// TwinCAT 3 PLC project PatchPress
// ProgramVersion: 3.1.4026.22
// libraries:
//   Tc2_Standard, * (Beckhoff Automation GmbH)
//   Tc2_System, * (Beckhoff Automation GmbH)
// project tree:
//   DUTs/01_Core/ E_CycleState.TcDUT, E_IndexFault.TcDUT, E_IndexState.TcDUT, E_InitialisingWaitReason.TcDUT, E_MachineState.TcDUT, E_MainDoorLockFault.TcDUT, E_MainDoorLockState.TcDUT, E_OperatorExchangeState.TcDUT, E_OperatorInstruction.TcDUT, E_PartDisposition.TcDUT (not stored), E_ProcessResultCode.TcDUT, E_StoppingWaitReason.TcDUT, E_TablePosition.TcDUT, ST_IndexStatus.TcDUT, ST_MachineCommand.TcDUT, ST_MachineConfig.TcDUT, ST_MachineInputs.TcDUT, ST_MachineOutputs.TcDUT, ST_MachinePermissives.TcDUT, ST_MachineStatus.TcDUT, ST_MainDoorLockStatus.TcDUT, ST_Nest.TcDUT, ST_NestStatistics.TcDUT, ST_OperatorStationStatus.TcDUT, ST_ProcessResult.TcDUT, ST_SafetyStatus.TcDUT (not stored), ST_TestHistory.TcDUT
//   DUTs/01_Core/Machine/ ST_PatchPressInputs.TcDUT, ST_PatchPressOutputs.TcDUT
//   DUTs/02_Components/Motion/ ST_Axis.TcDUT
//   DUTs/04_IO_Mapping/Terminals/ ST_EL3314.TcDUT, ST_EL6633.TcDUT, ST_EK1100.TcDUT (not stored), ST_EL1809.TcDUT (not stored), ST_EL1918.TcDUT, ST_EL2502.TcDUT, ST_EL2809.TcDUT (not stored), ST_EL2904.TcDUT, ST_EL3058.TcDUT, ST_EL3064.TcDUT, ST_EL6070.TcDUT (not stored), ST_EL6652.TcDUT (not stored), ST_EL6910.TcDUT, ST_EL7201.TcDUT, ST_EL9410.TcDUT (not stored), ST_Terminal_Info.TcDUT (not stored)
//   DUTs/07_HMI/ E_LEDs_Mode.TcDUT, E_PLC_Power.TcDUT (not stored), ST_HmiCommands.TcDUT, ST_HmiStatistics.TcDUT, ST_HmiStatus.TcDUT, ST_StatusBanner.TcDUT
//   DUTs/03_Stations/Common/ E_PatchPressStation.TcDUT, E_PatchStationState.TcDUT, ST_PatchStageStatus.TcDUT
//   DUTs/04_IO_Mapping/ ST_PhysicalInputs.TcDUT, ST_PhysicalOutputs.TcDUT
//   DUTs/05_AlarmsAndEvents/ E_AlarmId.TcDUT, E_AlarmSeverity.TcDUT, E_MachineAlarm.TcDUT, ST_ActiveAlarm.TcDUT (not stored), ST_ActiveEvents.TcDUT, ST_AlarmManagerStatus.TcDUT, ST_EVENT.TcDUT, ST_EventsAssigment.TcDUT, ST_EventsAssigmentGeneral.TcDUT (not stored), ST_EventsHistory.TcDUT (not stored), ST_StationEvents.TcDUT
//   GVLs/ GVL_Config.TcGVL, GVL_EtherCAT.TcGVL, GVL_HMI.TcGVL, GVL_IO.TcGVL (not stored), GVL_MASTER.TcGVL, GVL_Motion.TcGVL, GVL_PatchPress_Interface.TcGVL, GVL_Persistent.TcGVL, GVL_Safety.TcGVL
//   / PlcTask.TcTTO
//   POUs/00_Application/ PRG_HmiCommands.TcPOU, PRG_HmiStatus.TcPOU, PRG_Main.TcPOU, PRG_ReadInputs.TcPOU, PRG_WriteOutputs.TcPOU
//   POUs/01_Core/ I_ProcessEquipment.TcIO (not stored)
//   POUs/01_Core/Machine/ FB_IndexedPatchPressMachine.TcPOU, FB_PatchPressCommissioningGuard.TcPOU
//   POUs/01_Core/Process/ FB_ProcessCycle.TcPOU, FB_ProcessStation.TcPOU
//   POUs/02_Components/Door/ FB_MainDoorLock.TcPOU
//   POUs/02_Components/Index/ FB_IndexTable4.TcPOU, FB_NestTableManager.TcPOU, UINT_TO_E_TablePosition.TcPOU
//   POUs/02_Components/Pneumatics/ FB_PuckLocker.TcPOU, FB_Support.TcPOU
//   POUs/03_Stations/HeatStake/ FB_HeatStakeStation.TcPOU
//   POUs/03_Stations/Operator/ FB_OperatorStation.TcPOU
//   POUs/03_Stations/PatchDispense/ FB_PatchDispenseStation.TcPOU
//   POUs/03_Stations/Vision/ FB_VisionStation.TcPOU
//   POUs/04_IO_Mapping/ PRG_TerminalMapping.TcPOU
//   POUs/05_AlarmsAndEvents/ FB_EventsManager.TcPOU, PRG_Events.TcPOU
//   POUs/06_Utilities/ FB_TerminalInfo.TcPOU (not stored), F_ScaleLinear.TcPOU
//   POUs/ MAIN.TcPOU
// real-time tasks:
//   TASK PlcTask: cycle T#10ms, priority 20, ADS port 350
// motion (NC):
//   TASK NC-Task 1 SAF: cycle T#2ms, priority 4, ADS port 501
//   TASK NC-Task 1 SVB: cycle T#10ms, priority 8, ADS port 511
//   AXIS M1 (id 1)
//     OtherSettings: AllowMotionCmdToSlave=true
//     encoder EncType=19
//       EncPara: MaxCount=#xffffffff
//     drive DrvType=16
//       DrvPara: MaxCount=#xffffffff, DriveControlDWord=#x00020000
//         Analog: TorqueSetpointScale=10, ScaleFactorActTorque=0.1
//         TimeComp: TaskDelayCycles=1
//     controller CtrType=1
//       CtrPara: PriorControlFactor=1
//         Observer: BandWidth=20
//   AXIS M2 (id 2)
//     OtherSettings: AllowMotionCmdToSlave=true
//     encoder EncType=19
//       EncPara: MaxCount=#xffffffff
//     drive DrvType=16
//       DrvPara: MaxCount=#xffffffff, DriveControlDWord=#x00020000
//         Analog: TorqueSetpointScale=10, ScaleFactorActTorque=0.1
//         TimeComp: TaskDelayCycles=1
//     controller CtrType=1
//       CtrPara: PriorControlFactor=1
//         Observer: BandWidth=20
//   AXIS M3 (id 3)
//     OtherSettings: AllowMotionCmdToSlave=true
//     encoder EncType=19
//       EncPara: MaxCount=#xffffffff
//     drive DrvType=16
//       DrvPara: MaxCount=#xffffffff, DriveControlDWord=#x00020000
//         Analog: TorqueSetpointScale=10, ScaleFactorActTorque=0.1
//         TimeComp: TaskDelayCycles=1
//     controller CtrType=1
//       CtrPara: PriorControlFactor=1
//         Observer: BandWidth=20
// I/O:
//   DEVICE Device 1 (EtherCAT), AmsNetId 172.18.239.27.2.1
//     Term 1 (EK1100) [EK1100 EtherCAT Coupler (2A E-Bus)]
//       Term 2 (EL6070-0033) [EL6070-0033 1Ch. Licence key terminal, individual licences]
//       Term 3 (EL6910) [EL6910, TwinSAFE PLC]
//       Term 4 (EL1918) [EL1918, 8Ch. Safety Input 24V, TwinSAFE]
//         modules: Module 1 (FSOE), Module 2 (FSLOGIC)
//       Term 5 (EL1918) [EL1918, 8Ch. Safety Input 24V, TwinSAFE]
//         modules: Module 1 (FSOE), Module 2 (FSLOGIC)
//       Term 6 (EL2904) [EL2904, 4 Ch. Safety Output 24V, 0.5A, TwinSAFE]
//         modules: Module 1 (FSOES), Module 2 (DO)
//       Term 7 (EL1809) [EL1809 16Ch. Dig. Input 24V, 3ms]
//       Term 8 (EL1809) [EL1809 16Ch. Dig. Input 24V, 3ms]
//       Term 9 (EL2809-0015) [EL2809-0015 16Ch. Dig. Output 24V DC, 0.35A, not short-circuit proof]
//       Term 10 (EL2809-0015) [EL2809-0015 16Ch. Dig. Output 24V DC, 0.35A, not short-circuit proof]
//       Term 11 (EL3058) [EL3058 8Ch. Ana. Input 4-20mA]
//       Term 12 (EL9410) [EL9410 E-Bus Power Supplier  (Diagnostics)]
//       Term 13 (EL2502) [EL2502 2Ch. PWM output, 24V]
//       Term 14 (EL9576) [EL9576 Brake chopper terminal]
//       Term 15 (EL7201-9014) [EL7201-9014 1Ch. MDP742 Servo motor output stage with OCT (50V, 2.8A RMS) and STO input]
//       Term 16 (EL7201-9014) [EL7201-9014 1Ch. MDP742 Servo motor output stage with OCT (50V, 2.8A RMS) and STO input]
//       Term 17 (EL7201-9014) [EL7201-9014 1Ch. MDP742 Servo motor output stage with OCT (50V, 2.8A RMS) and STO input]
//       Term 18 (EL2904) [EL2904, 4 Ch. Safety Output 24V, 0.5A, TwinSAFE]
//         modules: Module 1 (FSOES), Module 2 (DO)
//       Term 19 (EL1809) [EL1809 16Ch. Dig. Input 24V, 3ms]
//       Term 20 (EL3314-0092) [EL3314-0092 4Ch. Ana Input Thermocouple (TC), TwinSAFE SC]
//       Term 21 (EL6633) [EL6633 PROFINET IO Controller]
//       Term 23 (EL9011) [EL9011 End Terminal]
//     Box 22 (VABX-A-S-EL-E12-CTED-ECM12) [VABX-A-S-EL-E12-CTED-ECM12] (disabled)
// variable links:
//   Device 1 (EtherCAT) <-> Device 1 (EtherCAT)/Term 1 (EK1100)/Term 3 (EL6910)
//     Term 1 (EK1100)/Term 18 (EL2904)/Module 1 (FSOES)/RxPDO/FSOE <-> ConnectionInputs/TwinSafeGroup1.Term 18 (EL2904) - Module 1 (FSOES)_6 TxPDO
//     Term 1 (EK1100)/Term 6 (EL2904)/Module 1 (FSOES)/RxPDO/FSOE <-> ConnectionInputs/TwinSafeGroup1.Term 6 (EL2904) - Module 1 (FSOES)_5 TxPDO
//     Term 1 (EK1100)/Term 18 (EL2904)/Module 1 (FSOES)/TxPDO/FSOE <-> ConnectionOutputs/TwinSafeGroup1.Term 18 (EL2904) - Module 1 (FSOES)_6 RxPDO
//     Term 1 (EK1100)/Term 6 (EL2904)/Module 1 (FSOES)/TxPDO/FSOE <-> ConnectionOutputs/TwinSafeGroup1.Term 6 (EL2904) - Module 1 (FSOES)_5 RxPDO
//     Term 1 (EK1100)/Term 4 (EL1918)/Module 1 (FSOE)/FSoE Inputs/FSOE <-> ConnectionOutputs/TwinSafeGroup1.Term 4 (EL1918) - Module 1 (FSOE)_3 RxPDO
//     Term 1 (EK1100)/Term 5 (EL1918)/Module 1 (FSOE)/FSoE Inputs/FSOE <-> ConnectionOutputs/TwinSafeGroup1.Term 5 (EL1918) - Module 1 (FSOE)_4 RxPDO
//     Term 1 (EK1100)/Term 4 (EL1918)/Module 1 (FSOE)/FSoE Outputs/FSOE <-> ConnectionInputs/TwinSafeGroup1.Term 4 (EL1918) - Module 1 (FSOE)_3 TxPDO
//     Term 1 (EK1100)/Term 5 (EL1918)/Module 1 (FSOE)/FSoE Outputs/FSOE <-> ConnectionInputs/TwinSafeGroup1.Term 5 (EL1918) - Module 1 (FSOE)_4 TxPDO
//   NC-Task 1 SAF/Axes/M1 <-> Device 1 (EtherCAT)/Term 1 (EK1100)/Term 15 (EL7201-9014)
//     Drive/Inputs/In/nDcOutputTime <-> InfoData/DcOutputShift
//     Drive/Inputs/In/nState1 <-> DRV Statusword/Statusword
//     Drive/Inputs/In/nState2 <-> DRV Statusword/Statusword @bit 8
//     Drive/Inputs/In/nState4 @bit 1 <-> WcState/InputToggle
//     Drive/Inputs/In/nState4 <-> WcState/WcState
//     Drive/Outputs/Out/nCtrl1 <-> DRV Controlword/Controlword
//     Drive/Outputs/Out/nCtrl2 <-> DRV Controlword/Controlword @bit 8
//     Drive/Outputs/Out/nDataOut2 <-> DRV Target velocity/Target velocity
//     Enc/Inputs/In/nDataIn1 <-> FB Position/Position
//     Enc/Inputs/In/nDcInputTime <-> InfoData/DcInputShift
//     Enc/Inputs/In/nState4 @bit 1 <-> WcState/InputToggle
//     Enc/Inputs/In/nState4 <-> WcState/WcState
//   NC-Task 1 SAF/Axes/M2 <-> Device 1 (EtherCAT)/Term 1 (EK1100)/Term 16 (EL7201-9014)
//     Drive/Inputs/In/nDcOutputTime <-> InfoData/DcOutputShift
//     Drive/Inputs/In/nState1 <-> DRV Statusword/Statusword
//     Drive/Inputs/In/nState2 <-> DRV Statusword/Statusword @bit 8
//     Drive/Inputs/In/nState4 @bit 1 <-> WcState/InputToggle
//     Drive/Inputs/In/nState4 <-> WcState/WcState
//     Drive/Outputs/Out/nCtrl1 <-> DRV Controlword/Controlword
//     Drive/Outputs/Out/nCtrl2 <-> DRV Controlword/Controlword @bit 8
//     Drive/Outputs/Out/nDataOut2 <-> DRV Target velocity/Target velocity
//     Enc/Inputs/In/nDataIn1 <-> FB Position/Position
//     Enc/Inputs/In/nDcInputTime <-> InfoData/DcInputShift
//     Enc/Inputs/In/nState4 @bit 1 <-> WcState/InputToggle
//     Enc/Inputs/In/nState4 <-> WcState/WcState
//   NC-Task 1 SAF/Axes/M3 <-> Device 1 (EtherCAT)/Term 1 (EK1100)/Term 17 (EL7201-9014)
//     Drive/Inputs/In/nDcOutputTime <-> InfoData/DcOutputShift
//     Drive/Inputs/In/nState1 <-> DRV Statusword/Statusword
//     Drive/Inputs/In/nState2 <-> DRV Statusword/Statusword @bit 8
//     Drive/Inputs/In/nState4 @bit 1 <-> WcState/InputToggle
//     Drive/Inputs/In/nState4 <-> WcState/WcState
//     Drive/Outputs/Out/nCtrl1 <-> DRV Controlword/Controlword
//     Drive/Outputs/Out/nCtrl2 <-> DRV Controlword/Controlword @bit 8
//     Drive/Outputs/Out/nDataOut2 <-> DRV Target velocity/Target velocity
//     Enc/Inputs/In/nDataIn1 <-> FB Position/Position
//     Enc/Inputs/In/nDcInputTime <-> InfoData/DcInputShift
//     Enc/Inputs/In/nState4 @bit 1 <-> WcState/InputToggle
//     Enc/Inputs/In/nState4 <-> WcState/WcState
//   PatchPress/PatchPress Instance <-> Device 1 (EtherCAT)/Term 1 (EK1100)/Term 10 (EL2809-0015)
//     PlcTask Inputs/GVL_EtherCAT.stTerm10_EL2809.stTerminalInfo.nTerminal_State <-> InfoData/State
//     PlcTask Outputs/GVL_EtherCAT.stTerm10_EL2809.iEL2809_Ch{1..16} <-> Channel {1..16}/Output  (16 links)
//   PatchPress/PatchPress Instance <-> Device 1 (EtherCAT)/Term 1 (EK1100)/Term 11 (EL3058)
//     PlcTask Inputs/GVL_EtherCAT.stTerm11_EL3058.iEL3058_Ch{1..8} <-> AI Standard Channel {1..8}/Value  (8 links)
//     PlcTask Inputs/GVL_EtherCAT.stTerm11_EL3058.stTerminalInfo.nTerminal_State <-> InfoData/State
//   PatchPress/PatchPress Instance <-> Device 1 (EtherCAT)/Term 1 (EK1100)/Term 19 (EL1809)
//     PlcTask Inputs/GVL_EtherCAT.stTerm19_EL1809.iEL1809_Ch{1..16} <-> Channel {1..16}/Input  (16 links)
//     PlcTask Inputs/GVL_EtherCAT.stTerm19_EL1809.stTerminalInfo.nTerminal_State <-> InfoData/State
//   PatchPress/PatchPress Instance <-> Device 1 (EtherCAT)/Term 1 (EK1100)/Term 3 (EL6910)
//     PlcTask Inputs/GVL_Safety.bMainDoorClosed <-> StandardInputs/Standard Out Var 8
//     PlcTask Inputs/GVL_Safety.bMainDoorLocked <-> StandardInputs/Standard Out Var 9
//     PlcTask Inputs/GVL_Safety.bMainDoorUnSafe <-> StandardInputs/Standard Out Var 10
//     PlcTask Inputs/GVL_Safety.bResetButtonPressed <-> StandardInputs/Standard Out Var 7
//     PlcTask Inputs/GVL_Safety.bSafetyOk <-> StandardInputs/Standard Out Var 12
//     PlcTask Inputs/GVL_Safety.bTwoHandSafe <-> StandardInputs/Standard Out Var 16
//     PlcTask Outputs/GVL_IO.stOutputs/bAirSupplyEnable <-> StandardOutputs/Standard In Var 11
//     PlcTask Outputs/GVL_IO.stOutputs/bMainDoorLockRequest <-> StandardOutputs/Standard In Var 14
//     PlcTask Outputs/GVL_IO.stOutputs/bSafetyErrorAcknowledgementRequest <-> StandardOutputs/Standard In Var 1
//     PlcTask Outputs/GVL_IO.stOutputs/bSafetyRunRequest <-> StandardOutputs/Standard In Var 15
//   PatchPress/PatchPress Instance <-> Device 1 (EtherCAT)/Term 1 (EK1100)/Term 7 (EL1809)
//     PlcTask Inputs/GVL_EtherCAT.stTerm7_EL1809.iEL1809_Ch{1..16} <-> Channel {1..16}/Input  (16 links)
//     PlcTask Inputs/GVL_EtherCAT.stTerm7_EL1809.stTerminalInfo.nTerminal_State <-> InfoData/State
//   PatchPress/PatchPress Instance <-> Device 1 (EtherCAT)/Term 1 (EK1100)/Term 8 (EL1809)
//     PlcTask Inputs/GVL_EtherCAT.stTerm8_EL1809.iEL1809_Ch{1..16} <-> Channel {1..16}/Input  (16 links)
//     PlcTask Inputs/GVL_EtherCAT.stTerm8_EL1809.stTerminalInfo.nTerminal_State <-> InfoData/State
//   PatchPress/PatchPress Instance <-> Device 1 (EtherCAT)/Term 1 (EK1100)/Term 9 (EL2809-0015)
//     PlcTask Inputs/GVL_EtherCAT.stTerm9_EL2809.stTerminalInfo.nTerminal_State <-> InfoData/State
//     PlcTask Outputs/GVL_EtherCAT.stTerm9_EL2809.iEL2809_Ch{1..16} <-> Channel {1..16}/Output  (16 links)

CONFIGURATION PatchPress
    RESOURCE PLC ON TwinCAT3
        TASK PlcTask(INTERVAL := T#10ms, PRIORITY := 20);
        PROGRAM MAIN WITH PlcTask : MAIN;
    END_RESOURCE
END_CONFIGURATION

// ---- DUTs/01_Core/E_CycleState.TcDUT
{attribute 'qualified_only'}
{attribute 'strict'}
{attribute 'to_string'}
TYPE E_CycleState :
(
    // CYCLE INITIALISATION
    Disabled                        := 0,
    Initialising                    := 10,
    WaitingForProcessCycleTrigger   := 20,
	
    // INDEX POSITION RECOVERY
    EvaluatingIndexPosition         := 30,
    RequestingIndexPositionRecovery := 40,
    WaitingForIndexPositionRecovery := 50,

    // INDEX MOVEMENT
    ValidatingIndexPermissives      := 60,
    RequestingIndexMove             := 70,
    WaitingForIndexStart            := 80,
    WaitingForIndexComplete         := 90,

    // NEST AND PROCESS PREPARATION
    UpdatingNestPositions           := 100,
    EvaluatingProcessNest           := 110,
    SkippingProcessNest             := 120,

    // SUPPORT EXTENSION
    RequestingSupportsExtend        := 130,
    WaitingForSupportsExtended      := 140,

    // PROCESS EXECUTION
    PreparingProcessStations        := 150,
    WaitingForProcessStationsReady  := 160,
    StartingProcesses               := 170,
    WaitingForProcessesRunning      := 180,
    WaitingForProcessesComplete     := 190,

    // PROCESS RESULT
    CapturingProcessResult          := 200,
    StoringProcessResult            := 210,

    // SUPPORT RETRACTION
    RequestingSupportsRetract       := 220,
    WaitingForSupportsRetracted     := 230,

    // OPERATOR EXCHANGE
    PreparingOperatorExchange       := 240,
    WaitingForOperatorExchange      := 250,
    ConfirmingOperatorExchange      := 260,

    // CYCLE COMPLETION
    CycleComplete                   := 270,

    // TERMINAL STATES
    ControlledStop                  := 900,
    Fault                           := 999
);
END_TYPE

// ---- DUTs/01_Core/E_IndexFault.TcDUT
{attribute 'qualified_only'}
{attribute 'strict'}
{attribute 'to_string'}
TYPE E_IndexFault :
(
    None := 0,
    InitialPositionInvalid,
    SupportRetractTimeout,
    RotationTimeout,
    StopAndLockTimeout,
    PositionInvalid,
    SupportExtendTimeout,
    TwoHandReleasedDuringMovement,
    WrongPositionTimeout,
    SafetyLostDuringMovement,
    MovementPermissiveLost
);
END_TYPE

// ---- DUTs/01_Core/E_IndexState.TcDUT
{attribute 'qualified_only'}
{attribute 'strict'}
{attribute 'to_string'}
TYPE E_IndexState :
(
    Disabled := 0,
    Initialising,
    Idle,
    RetractingSupport,
    WaitingSupportRetracted,
    RotatingPortA,
    WrongPositionRecovery,
    StoppingPortB,
    VerifyingPosition,
    ExtendingSupport,
    WaitingSupportExtended,
    ProcessPositionReady,
    WaitingOperatorExchange,
    Complete,
    Stopping,
    Fault
);
END_TYPE

// ---- DUTs/01_Core/E_InitialisingWaitReason.TcDUT
{attribute 'qualified_only'}
{attribute 'strict'}
{attribute 'to_string'}
TYPE E_InitialisingWaitReason :
(
    None := 0,
    SafetyNotReady := 10,
    FsoeNotReady := 20,
    SafetyLogicNotReady := 30,
    AirSupplyNotReady := 40,
    MainDoorNotReady := 50,
    IndexNotReady := 60,
    StationsNotHome := 70
);
END_TYPE

// ---- DUTs/01_Core/E_MachineState.TcDUT
{attribute 'qualified_only'}
{attribute 'strict'}
{attribute 'to_string'}
TYPE E_MachineState :
(
    PowerUp      := 0,
    Fault        := 1,
    Stopping     := 2,
    Stopped      := 3,
    Initialising := 4,
    ReadyToStart := 5,
    AutoCycle    := 6,
    Manual       := 7
);
END_TYPE

// ---- DUTs/01_Core/E_MainDoorLockFault.TcDUT
{attribute 'qualified_only'}
{attribute 'strict'}
{attribute 'to_string'}
TYPE E_MainDoorLockFault :
(
    None := 0,
    LockTimeout := 10,
    UnlockTimeout := 20,
    DoorNotClosed := 30,
    FeedbackMismatch := 40
);
END_TYPE

// ---- DUTs/01_Core/E_MainDoorLockState.TcDUT
{attribute 'qualified_only'}
{attribute 'strict'}
{attribute 'to_string'}
TYPE E_MainDoorLockState :
(
    Disabled := 0,
    Unlocked := 10,
    Locking := 20,
    Locked := 30,
    Unlocking := 40,
    Fault := 999
);
END_TYPE

// ---- DUTs/01_Core/E_OperatorExchangeState.TcDUT
{attribute 'qualified_only'}
{attribute 'strict'}
{attribute 'to_string'}
TYPE E_OperatorExchangeState :
(
    Idle := 0,
    EvaluateNest := 10,
    WaitingForPartRemoval := 20,
    WaitingForRejectConfirmation := 30,
    WaitingForPuckRemoval := 40,
    WaitingForNewPuck := 50,
    WaitingForPuckLocked := 60,
    WaitingForPartLoading := 70,
    ExchangeComplete := 80,
    WaitingForTableIndexComplete := 90,
    Fault := 999
);
END_TYPE

// ---- DUTs/01_Core/E_OperatorInstruction.TcDUT
{attribute 'qualified_only'}
{attribute 'strict'}
{attribute 'to_string'}
TYPE E_OperatorInstruction :
(
    None := 0,
    LoadInitialPuck := 10,
    WaitPuckLocking := 20,
    RemovePassedPart := 30,
    RemoveFailedPart := 40,
    PlacePartInRejectBin := 50,
    RemoveReleasedPuck := 60,
    LoadNewPuck := 70,
    LoadPart := 80,
    ReadyToIndex := 90,
    ReadyToIndexEmpty := 100,
    TableIndexing := 110,
    RestoreUnexpectedlyRemovedPuck := 120
);
END_TYPE

// ---- DUTs/01_Core/E_ProcessResultCode.TcDUT
{attribute 'qualified_only'}
{attribute 'strict'}
{attribute 'to_string'}
TYPE E_ProcessResultCode :
(
	None := 0,
    Pass,
    Fail,
    Aborted,
    EquipmentFault,
    CommunicationFault,
    Timeout
);
END_TYPE

// ---- DUTs/01_Core/E_StoppingWaitReason.TcDUT
{attribute 'qualified_only'}
{attribute 'strict'}
{attribute 'to_string'}
TYPE E_StoppingWaitReason :
(
    None := 0,
    IndexStillMoving := 10,
    MainDoorTransition := 20
);
END_TYPE

// ---- DUTs/01_Core/E_TablePosition.TcDUT
{attribute 'qualified_only'}
{attribute 'strict'}
{attribute 'to_string'}
TYPE E_TablePosition :
(
	Unknown := 0,
    Position1 := 1,
    Position2 := 2,
    Position3 := 3,
    Position4 := 4
);
END_TYPE

// ---- DUTs/01_Core/Machine/ST_PatchPressInputs.TcDUT
TYPE ST_PatchPressInputs :
STRUCT
    // EPLAN Term 7 - EL1809
    b48VPowerSupplyOk                   : BOOL;
    bLoadingStationEaglePresent         : BOOL;
    bRejectChutePartPresent             : BOOL;
    bHeatStakeEagleAssemblyPresent      : BOOL;
    bHeatStakePatchPresent              : BOOL;
    bPbupMagnetPresent                  : BOOL;

    // EPLAN Term 8 - EL1809
    bStation1SupportRetracted           : BOOL;
    bStation1SupportExtended            : BOOL;
    bStation2SupportRetracted           : BOOL;
    bStation2SupportExtended            : BOOL;
    bStation3SupportRetracted           : BOOL;
    bStation3SupportExtended            : BOOL;
    bHorizontalMiniSlideRetracted       : BOOL;
    bHorizontalMiniSlideExtended        : BOOL;
    bVerticalMiniSlideRetracted         : BOOL;
    bVerticalMiniSlideExtended          : BOOL;
    bIntermediateModuleRetracted        : BOOL;
    bIntermediateModuleExtended         : BOOL;
    bRotaryGripperOpened                : BOOL;
    bRotaryGripperClosed                : BOOL;
    bRotaryGripperPick0                 : BOOL;
    bRotaryGripperPlace180              : BOOL;

    // EPLAN Term 19 - EL1809
    bMembraneTransferRetracted          : BOOL;
    bMembraneTransferExtended           : BOOL;
    bMiddleRockerDown                   : BOOL;
    bMiddleRockerUp                     : BOOL;
    bBottomRockerDown                   : BOOL;
    bBottomRockerUp                     : BOOL;
    bTopRockerDown                      : BOOL;
    bTopRockerUp                        : BOOL;

    // EPLAN Term 11 / 20
    iMainAirPressureRaw                 : INT;
    iProportionalPressureActualRaw      : INT;
    iCartridgeHeater1TemperatureRaw     : INT;
    iCartridgeHeater2TemperatureRaw     : INT;
    iOverTemperatureRaw                 : INT;
END_STRUCT
END_TYPE

// ---- DUTs/01_Core/Machine/ST_PatchPressOutputs.TcDUT
TYPE ST_PatchPressOutputs :
STRUCT
    // Pneumatic commands are logical commands only at this stage.
    // Physical Festo manifold PDO mapping must be created after the manifold scan.
    bStation1SupportExtend              : BOOL;
    bStation1SupportRetract             : BOOL;
    bStation2SupportExtend              : BOOL;
    bStation2SupportRetract             : BOOL;
    bStation3SupportExtend              : BOOL;
    bStation3SupportRetract             : BOOL;
    bHorizontalMiniSlideExtend          : BOOL;
    bHorizontalMiniSlideRetract         : BOOL;
    bVerticalMiniSlideExtend            : BOOL;
    bVerticalMiniSlideRetract           : BOOL;
    bIntermediateModuleExtend           : BOOL;
    bIntermediateModuleRetract          : BOOL;
    bRotaryGripperOpen                  : BOOL;
    bRotaryGripperClose                 : BOOL;
    bRotaryGripperPick0                 : BOOL;
    bRotaryGripperPlace180              : BOOL;
    bMembraneTransferExtend             : BOOL;
    bMembraneTransferRetract            : BOOL;
    bMiddleRockerDown                   : BOOL;
    bMiddleRockerUp                     : BOOL;
    bBottomRockerDown                   : BOOL;
    bBottomRockerUp                     : BOOL;
    bTopRockerDown                      : BOOL;
    bTopRockerUp                        : BOOL;

    // Heater / pressure logical commands.
    rHeater1DutyPercent                 : REAL;
    rHeater2DutyPercent                 : REAL;
    rPressureSetpointBar                : REAL;
END_STRUCT
END_TYPE

// ---- DUTs/01_Core/ST_IndexStatus.TcDUT
TYPE ST_IndexStatus :
STRUCT
    eState                    : E_IndexState;
    eFault                    : E_IndexFault;
    eCurrentPosition          : E_TablePosition;

    bReady                    : BOOL;
    bBusy                     : BOOL;
    bFaulted                  : BOOL;
    bDonePulse                : BOOL;

    bManualMoveActive         : BOOL;
    bPositionRecoveryActive   : BOOL;
    bSamePositionDetected     : BOOL;
    bWrongPositionTimerActive : BOOL;
    bTwoHandRequired          : BOOL;

    bProcessPositionReady     : BOOL;
    bWaitingOperatorExchange  : BOOL;

    bSupportRetracted         : BOOL;
    bSupportExtended          : BOOL;
    bTableReady               : BOOL;
    bTableLocked              : BOOL;
	
END_STRUCT
END_TYPE

// ---- DUTs/01_Core/ST_MachineCommand.TcDUT
TYPE ST_MachineCommand :
STRUCT
    bStart                : BOOL;
    bStop                 : BOOL;
    bReset                : BOOL;
    bManualRequest        : BOOL;
    bManualIndexForward   : BOOL;
    bManualIndexHome      : BOOL;
    bIndexerManualEnable  : BOOL;
    bManualMainDoorUnlock : BOOL;
    bAcknowledge          : BOOL;
    bAcknowledgePuckRemovalFault : BOOL;
    uiResetStatisticsNestId : UINT;
END_STRUCT
END_TYPE

// ---- DUTs/01_Core/ST_MachineConfig.TcDUT
TYPE ST_MachineConfig :
STRUCT
    tInitialiseTimeout       : TIME := T#20S;
    tStoppingTimeout         : TIME := T#15S;
    tIndexTimeout            : TIME := T#10S;
    tIndexRotateDelay        : TIME := T#500MS;
    tIndexStopDelay          : TIME := T#1S;
    tIndexSupportTimeout     : TIME := T#5S;
    tTwoHandHold             : TIME := T#500MS;
    tTwoHandRecoveryTimeout  : TIME := T#10S;
    tDoorLockTimeout         : TIME := T#10S;
    tDoorUnlockTimeout       : TIME := T#10S;
    tOperatorIdleTimeout     : TIME := T#30S;
    eOperatorPosition        : E_TablePosition := E_TablePosition.Position1;
    ePatchDispensePosition   : E_TablePosition := E_TablePosition.Position2;
    eHeatStakePosition       : E_TablePosition := E_TablePosition.Position3;
    eVisionPosition          : E_TablePosition := E_TablePosition.Position4;
    eRejectPosition          : E_TablePosition := E_TablePosition.Position1;
    bRequireTwoHandsForIndex : BOOL := TRUE;
    bAllowEmptyNestIndex     : BOOL := TRUE;
    bRequireRejectConfirm    : BOOL := TRUE;
    aNestEnabled             : ARRAY[1..4] OF BOOL := [TRUE, TRUE, TRUE, TRUE];
END_STRUCT
END_TYPE

// ---- DUTs/01_Core/ST_MachineInputs.TcDUT
TYPE ST_MachineInputs :
STRUCT
    bStartButton                  : BOOL;
    bStopButton                   : BOOL;
    bResetButton                  : BOOL;
    bTwoHandsSafe                 : BOOL;
    bTouchButtonLeft              : BOOL;
    bTouchButtonRight             : BOOL;
    bUp24VPowerSupplyOk           : BOOL;
    bUs24VPowerSupplyOk           : BOOL;
    b48VPowerSupplyOk             : BOOL;
    bEmergencyStopChannel1        : BOOL;
    bEmergencyStopChannel2        : BOOL;
    bMainDoorChannel1             : BOOL;
    bMainDoorChannel2             : BOOL;
    bMainDoorFeedback             : BOOL;
    bLeftFlapChannel1             : BOOL;
    bLeftFlapChannel2             : BOOL;
    bRightFlapChannel1            : BOOL;
    bRightFlapChannel2            : BOOL;
    bMainDoorClosed               : BOOL;
    bMainDoorLocked               : BOOL;
    bMainDoorUnsafe               : BOOL;
    bMainDoorDiagnosticOk         : BOOL;
    bMs6FeedbackOk                : BOOL;
    bAirExhausted                 : BOOL;
    stSafety                      : ST_SafetyStatus;
    bEventFault                   : BOOL;
    bEventCycleStopRequest        : BOOL;
    bIndexReady                   : BOOL;
    bIndexLocked                  : BOOL;
    bIndexCompletedSensor         : BOOL;
    eIndexPosition                : E_TablePosition;
    bLoadingStationEaglePresent   : BOOL;
    bRejectChutePartPresent       : BOOL;
    bHeatStakeEaglePresent        : BOOL;
    bHeatStakePatchPresent        : BOOL;
    bPbupMagnetPresent            : BOOL;
    bStation1SupportRetracted     : BOOL;
    bStation1SupportExtended      : BOOL;
    bStation2SupportRetracted     : BOOL;
    bStation2SupportExtended      : BOOL;
    bStation3SupportRetracted     : BOOL;
    bStation3SupportExtended      : BOOL;
    bHorizontalMiniSlideRetracted : BOOL;
    bHorizontalMiniSlideExtended  : BOOL;
    bVerticalMiniSlideRetracted   : BOOL;
    bVerticalMiniSlideExtended    : BOOL;
    bIntermediateModuleRetracted  : BOOL;
    bIntermediateModuleExtended   : BOOL;
    bRotaryGripperOpened          : BOOL;
    bRotaryGripperClosed          : BOOL;
    bRotaryGripperPick0           : BOOL;
    bRotaryGripperPlace180        : BOOL;
    bMembraneTransferRetracted    : BOOL;
    bMembraneTransferExtended     : BOOL;
    bMiddleRockerDown             : BOOL;
    bMiddleRockerUp               : BOOL;
    bBottomRockerDown             : BOOL;
    bBottomRockerUp               : BOOL;
    bTopRockerDown                : BOOL;
    bTopRockerUp                  : BOOL;
    uiMainAirPressureRaw          : UINT;
    uiPressureRegulatorActualRaw  : UINT;
END_STRUCT
END_TYPE

// ---- DUTs/01_Core/ST_MachineOutputs.TcDUT
TYPE ST_MachineOutputs :
STRUCT
    bSafetyRunRequest                  : BOOL;
    bSafetyResetRequest                : BOOL;
    bSafetyErrorAcknowledgementRequest : BOOL;
    bAirSupplyEnable                   : BOOL;
    bMainDoorLockRequest               : BOOL;
    bIndexRotatePortA                  : BOOL;
    bIndexStopPortB                    : BOOL;
    bIndexSupportExtend                : BOOL;
    bIndexSupportRetract               : BOOL;
    bLedStart                          : BOOL;
    bLedReset                          : BOOL;
    bLedPass                           : BOOL;
    bLedFail                           : BOOL;
    bInternalLight                     : BOOL;
    bNestLight                         : BOOL;
END_STRUCT
END_TYPE

// ---- DUTs/01_Core/ST_MachinePermissives.TcDUT
TYPE ST_MachinePermissives :
STRUCT
    bSafetyIndexPermissive   : BOOL;
    bOperatorIndexPermissive : BOOL;
    bStationsIndexPermissive : BOOL;
    bIndexMoveAllowed        : BOOL;
    bAirSupplyReady          : BOOL;
    bDoorInitialisationReady : BOOL;
    bIndexInitialisationReady: BOOL;
    bStationsHome            : BOOL;
    bInitialisationAllowed   : BOOL;
    bAutoCycleAllowed        : BOOL;
END_STRUCT
END_TYPE

// ---- DUTs/01_Core/ST_MachineStatus.TcDUT
TYPE ST_MachineStatus :
STRUCT
    eMachineState           : E_MachineState;
    eIndexState             : E_IndexState;
    stIndexStatus           : ST_IndexStatus;
    stMainDoorLock          : ST_MainDoorLockStatus;
    eInitialisingWaitReason : E_InitialisingWaitReason;
    eStoppingWaitReason     : E_StoppingWaitReason;
    eOperatorExchangeState  : E_OperatorExchangeState;
    eOperatorInstruction    : E_OperatorInstruction;
    stOperatorStation       : ST_OperatorStationStatus;
    stPatchDispense         : ST_PatchStageStatus;
    stHeatStake             : ST_PatchStageStatus;
    stVision                : ST_PatchStageStatus;
    bReady                  : BOOL;
    bBusy                   : BOOL;
    bFaulted                : BOOL;
    bInitialisationTimeoutFault : BOOL;
    bStoppingTimeoutFault   : BOOL;
    bSafetyStopRequested    : BOOL;
    bSafetyRunRequested     : BOOL;
    bEventFault             : BOOL;
    bCycleStopRequested     : BOOL;
    bIndexPermissive        : BOOL;
    bEnableSetting          : BOOL;
    bAllStationsCommissioned: BOOL;
    bAutoCycleAllowed       : BOOL;
    stPermissives           : ST_MachinePermissives;
    stLastResult            : ST_ProcessResult;
    aNest                   : ARRAY[1..4] OF ST_Nest;
    aNestStatistics         : ARRAY[1..4] OF ST_NestStatistics;
    sMachineMessage         : STRING(160);
    sOperatorMessage        : STRING(255);
    sAutoCycleBlockReason   : STRING(160);
END_STRUCT
END_TYPE

// ---- DUTs/01_Core/ST_MainDoorLockStatus.TcDUT
TYPE ST_MainDoorLockStatus :
STRUCT
    eState                  : E_MainDoorLockState;
    eFault                  : E_MainDoorLockFault;
    bDoorClosed             : BOOL;
    bDoorLocked             : BOOL;
    bDoorUnsafe             : BOOL;
    bLockRequest            : BOOL;
    bLockOutput             : BOOL;
    bReadyForAutomatic      : BOOL;
    bUnlockPermissive       : BOOL;
    bFaulted                : BOOL;
    sMessage                : STRING(160);
END_STRUCT
END_TYPE

// ---- DUTs/01_Core/ST_Nest.TcDUT
TYPE ST_Nest :
STRUCT
    nId                       : UINT;
    ePosition                 : E_TablePosition;
    bEnabled                  : BOOL;
    bPartPresent              : BOOL;
    bPreviousPartPresent      : BOOL;
    bPartLoadedPulse          : BOOL;
    bPartRemovedPulse         : BOOL;
    bProcessRequired          : BOOL;
    bProcessComplete          : BOOL;
    eDisposition              : E_PartDisposition;
    bDispositionSent          : BOOL;
    bOperatorExchangeComplete : BOOL;
    stPatchDispenseResult     : ST_ProcessResult;
    stHeatStakeResult         : ST_ProcessResult;
    stVisionResult            : ST_ProcessResult;
    stResult                  : ST_ProcessResult;
    bStatisticsCounted        : BOOL;
END_STRUCT
END_TYPE

// ---- DUTs/01_Core/ST_NestStatistics.TcDUT
TYPE ST_NestStatistics :
STRUCT
    uiNestId       : UINT;
    udiTotalTests  : UDINT;
    udiGoodParts   : UDINT;
    udiBadParts    : UDINT;
    lrEfficiency   : LREAL;
END_STRUCT
END_TYPE

// ---- DUTs/01_Core/ST_OperatorStationStatus.TcDUT
TYPE ST_OperatorStationStatus :
STRUCT
    eState                  : E_OperatorExchangeState;
    eInstruction            : E_OperatorInstruction;
    bExchangeComplete       : BOOL;
    bIndexPermissive        : BOOL;
    bPartRemovedConfirmed   : BOOL;
    bRejectConfirmed        : BOOL;
    bRejectArmed            : BOOL;
    bRejectEdgeAccepted     : BOOL;
    bRejectWaitingForClear  : BOOL;
    bPartPresent            : BOOL;
    bRejectChutePartPresent : BOOL;
    bResultValid            : BOOL;
    bResultPassed           : BOOL;
    sMessage                : STRING(255);
END_STRUCT
END_TYPE

// ---- DUTs/01_Core/ST_ProcessResult.TcDUT
TYPE ST_ProcessResult :
STRUCT
	bValid          : BOOL;
    bPassed         : BOOL;
    eCode           : E_ProcessResultCode;
    udiFaultCode    : UDINT;
    udiAlertCode    : UDINT;
    usiRecipe       : USINT;
    lrDispenseValue : LREAL;
    sDetail         : STRING(120);
END_STRUCT
END_TYPE

// ---- DUTs/01_Core/ST_TestHistory.TcDUT
TYPE ST_TestHistory :
STRUCT
    uiNestId            : UINT;
    eResult             : E_PartDisposition;
    bPatchDispenseValid : BOOL;
    bPatchDispensePass  : BOOL;
    bHeatStakeValid     : BOOL;
    bHeatStakePass      : BOOL;
    bVisionValid        : BOOL;
    bVisionPass         : BOOL;
    sResult             : STRING(20);
    sPatchDispenseResult: STRING(20);
    sHeatStakeResult    : STRING(20);
    sVisionResult       : STRING(20);
    sTime               : STRING(255);
    sDate               : STRING(255);
END_STRUCT
END_TYPE

// ---- DUTs/02_Components/Motion/ST_Axis.TcDUT
TYPE ST_Axis :
STRUCT
    // TwinCAT NC axis reference. Link this member to the corresponding NC axis.
    Axis                : AXIS_REF;

    // Standardised application-facing axis status / diagnostics.
    // These members may be linked to NC values directly during commissioning,
    // or populated later by the common motion component FB.
    bEnabled            : BOOL;
    bOperational        : BOOL;
    bHomed              : BOOL;
    bMoving             : BOOL;
    bStandstill         : BOOL;
    bError              : BOOL;

    lrActPosition       : LREAL;
    lrActVelocity       : LREAL;
    lrActTorque         : LREAL;

    udiErrorId          : UDINT;
END_STRUCT
END_TYPE

// ---- DUTs/04_IO_Mapping/Terminals/ST_EL3314.TcDUT
TYPE ST_EL3314 :
STRUCT
 
	//--------------------------------------------------------------------------------------------------------
	sTerminalName                                           :   STRING(200):= 'EL3314-0092 | 4-channel Analog Input, Thermocouple, TwinSAFE SC';
    //============================================================================================================================	
	// TERMINAL - EL3314-0092 | 4-channel Analog Input, Thermocouple, TwinSAFE SC (Term 20)	
	iEL3314_Ch1               				AT %I*			: 	DINT;	// EL3314 channel 1
	iEL3314_Ch2                   			AT %I*			: 	DINT;	// EL3314 channel 2
	iEL3314_Ch3        						AT %I*	 		: 	DINT;	// EL3314 channel 3
	iEL3314_Ch4	   							AT %I*	 		: 	DINT;	// EL3314 channel 4

	stTerminalInfo											: 	ST_Terminal_Info;	

END_STRUCT
END_TYPE

// ---- DUTs/04_IO_Mapping/Terminals/ST_EL6633.TcDUT
TYPE ST_EL6633 :
STRUCT
	sTerminalName : STRING(80) := 'EL6633 | 2-Port PROFINET Communication Interface';

    stTerminalInfo : ST_Terminal_Info;
END_STRUCT
END_TYPE

// ---- DUTs/07_HMI/E_LEDs_Mode.TcDUT
{attribute 'qualified_only'}
{attribute 'strict'}
{attribute 'to_string'}
TYPE E_LEDs_Mode :
(
    OFF := 0,
    ON := 1,
    FLASHING := 2
);
END_TYPE

// ---- DUTs/07_HMI/ST_HmiCommands.TcDUT
TYPE ST_HmiCommands :
STRUCT
    bStart                 : BOOL;
    bStop                  : BOOL;
    bReset                 : BOOL;
    bAcknowledge           : BOOL;
    bManualRequest         : BOOL;
    bIndexerManualEnable   : BOOL;
    bManualIndexForward    : BOOL;
    bManualIndexHome       : BOOL;
    bManualMainDoorUnlock  : BOOL;
    uiResetStatisticsNestId: UINT;
END_STRUCT
END_TYPE

// ---- DUTs/07_HMI/ST_HmiStatistics.TcDUT
TYPE ST_HmiStatistics :
STRUCT
    // OVERALL PRODUCTION
    udiTotalCycles          : UDINT;
    udiTotalPass            : UDINT;
    udiTotalFail            : UDINT;

    // PER-NEST PRODUCTION
    aNest                   : ARRAY[1..4] OF ST_NestStatistics;

    // MACHINE STATISTICS
    udiEquipmentFaults      : UDINT;
    udiIndexFaults          : UDINT;
    udiSafetyStops          : UDINT;
    udiAbortedCycles        : UDINT;

    dtLastCycleCompleted    : DATE_AND_TIME;
END_STRUCT
END_TYPE

// ---- DUTs/07_HMI/ST_HmiStatus.TcDUT
TYPE ST_HmiStatus :
STRUCT
    eMachineState             : E_MachineState;
    eIndexState               : E_IndexState;
    eIndexPosition            : E_TablePosition;
    iNestRotationAngle        : INT;
    bReady                    : BOOL;
    bBusy                     : BOOL;
    bFaulted                  : BOOL;
    bTwoHandsSafe             : BOOL;
    bLoadingStationEaglePresent : BOOL;
    bRejectChutePartPresent   : BOOL;
    bHeatStakeEaglePresent    : BOOL;
    bHeatStakePatchPresent    : BOOL;
    bPbupMagnetPresent        : BOOL;
    bIndexReady               : BOOL;
    bIndexLocked              : BOOL;
    bIndexCompletedSensor     : BOOL;
    bMainDoorClosed           : BOOL;
    bMainDoorLocked           : BOOL;
    bStartButtonActive        : BOOL;
    bStopButtonActive         : BOOL;
    bResetButtonActive        : BOOL;
    bStartButtonLamp          : BOOL;
    bUp24VPowerSupplyOk       : BOOL;
    bUs24VPowerSupplyOk       : BOOL;
    b48VPowerSupplyOk         : BOOL;
    bMainDoorDiagnosticOk     : BOOL;
    bMs6FeedbackOk            : BOOL;
    bAirExhausted             : BOOL;
    bLeftFlapSafe             : BOOL;
    bRightFlapSafe            : BOOL;
    bEnableSettings           : BOOL;
    bAllStationsCommissioned  : BOOL;
    bAutoCycleAllowed         : BOOL;
    stPatchDispense           : ST_PatchStageStatus;
    stHeatStake               : ST_PatchStageStatus;
    stVision                  : ST_PatchStageStatus;
    eOperatorInstruction      : E_OperatorInstruction;
    stOperatorStation         : ST_OperatorStationStatus;
    aNest                     : ARRAY[1..4] OF ST_Nest;
    sMachineMessage           : STRING(160);
    sOperatorMessage          : STRING(255);
    sAutoCycleBlockReason     : STRING(160);
END_STRUCT
END_TYPE

// ---- DUTs/07_HMI/ST_StatusBanner.TcDUT
TYPE ST_StatusBanner :
STRUCT
    sMachineStatusText : STRING(80);
    sBannerBckColor    : STRING(40);
    sBannerTextColor   : STRING(40);
END_STRUCT
END_TYPE

// ---- DUTs/03_Stations/Common/E_PatchPressStation.TcDUT
{attribute 'qualified_only'}
{attribute 'strict'}
{attribute 'to_string'}
TYPE E_PatchPressStation :
(
    Unknown := 0,
    Operator := 1,
    PatchDispense := 2,
    HeatStake := 3,
    Vision := 4
);
END_TYPE

// ---- DUTs/03_Stations/Common/E_PatchStationState.TcDUT
{attribute 'qualified_only'}
{attribute 'strict'}
{attribute 'to_string'}
TYPE E_PatchStationState :
(
    Disabled := 0,
    Homing := 10,
    Ready := 20,
    Processing := 30,
    Complete := 40,
    Fault := 100
);
END_TYPE

// ---- DUTs/03_Stations/Common/ST_PatchStageStatus.TcDUT
TYPE ST_PatchStageStatus :
STRUCT
    eState              : E_PatchStationState;
    bCommissioned       : BOOL;
    bHome               : BOOL;
    bReady              : BOOL;
    bBusy               : BOOL;
    bComplete           : BOOL;
    bFault              : BOOL;
    bPartPresent        : BOOL;
    sDiagnostic         : STRING(120);
END_STRUCT
END_TYPE

// ---- DUTs/04_IO_Mapping/ST_PhysicalInputs.TcDUT
TYPE ST_PhysicalInputs :
STRUCT
    bEmergencyStopChannel1 : BOOL;
    bEmergencyStopChannel2 : BOOL;
    bResetButton           : BOOL;
    bMainDoorChannel1      : BOOL;
    bMainDoorChannel2      : BOOL;
    bMainDoorFeedback      : BOOL;
    bMs6FeedbackOk         : BOOL;
    bAirExhausted          : BOOL;
    bTouchButtonLeft       : BOOL;
    bTouchButtonRight      : BOOL;
    bRightFlapChannel1     : BOOL;
    bRightFlapChannel2     : BOOL;
    bLeftFlapChannel1      : BOOL;
    bLeftFlapChannel2      : BOOL;
    bStartButton           : BOOL;
    bStopButton            : BOOL;
    bUp24VPowerSupplyOk    : BOOL;
    bUs24VPowerSupplyOk    : BOOL;
    b48VPowerSupplyOk      : BOOL;
    bIndexPositionSensor1  : BOOL;
    bIndexPositionSensor2  : BOOL;
    bIndexPositionSensor3  : BOOL;
    bIndexCompletedSensor  : BOOL;
    bIndexLocked           : BOOL;
    bIndexReady            : BOOL;
    eIndexPosition         : E_TablePosition;
    bLoadingStationEaglePresent : BOOL;
    bRejectChutePartPresent : BOOL;
    bHeatStakeEaglePresent : BOOL;
    bHeatStakePatchPresent : BOOL;
    bPbupMagnetPresent     : BOOL;
    bStation1SupportRetracted : BOOL;
    bStation1SupportExtended  : BOOL;
    bStation2SupportRetracted : BOOL;
    bStation2SupportExtended  : BOOL;
    bStation3SupportRetracted : BOOL;
    bStation3SupportExtended  : BOOL;
    bHorizontalMiniSlideRetracted : BOOL;
    bHorizontalMiniSlideExtended  : BOOL;
    bVerticalMiniSlideRetracted : BOOL;
    bVerticalMiniSlideExtended : BOOL;
    bIntermediateModuleRetracted : BOOL;
    bIntermediateModuleExtended : BOOL;
    bRotaryGripperOpened : BOOL;
    bRotaryGripperClosed : BOOL;
    bRotaryGripperPick0 : BOOL;
    bRotaryGripperPlace180 : BOOL;
    bMembraneTransferRetracted : BOOL;
    bMembraneTransferExtended : BOOL;
    bMiddleRockerDown : BOOL;
    bMiddleRockerUp : BOOL;
    bBottomRockerDown : BOOL;
    bBottomRockerUp : BOOL;
    bTopRockerDown : BOOL;
    bTopRockerUp : BOOL;
    uiMainAirPressureRaw : UINT;
    uiPressureRegulatorActualRaw : UINT;
    bSafetyOk : BOOL;
    bMainDoorClosed : BOOL;
    bMainDoorLocked : BOOL;
    bMainDoorUnsafe : BOOL;
    bMainDoorDiagnosticOk : BOOL;
    bTwoHandsSafe : BOOL;
END_STRUCT
END_TYPE

// ---- DUTs/04_IO_Mapping/ST_PhysicalOutputs.TcDUT
TYPE ST_PhysicalOutputs :
STRUCT
    bSafetyRunRequest                  : BOOL;
    bSafetyResetRequest                : BOOL;
    bSafetyErrorAcknowledgementRequest : BOOL;
    bAirSupplyEnable                   : BOOL;
    bMainDoorLockRequest               : BOOL;
    bIndexRotatePortA                  : BOOL;
    bIndexStopPortB                    : BOOL;
    bLedStart                          : BOOL;
    bLedReset                          : BOOL;
    bStatusIndicator                  : BOOL;
    bInternalLight                    : BOOL;
    bNestLight                        : BOOL;
END_STRUCT
END_TYPE

// ---- DUTs/04_IO_Mapping/Terminals/ST_EL1918.TcDUT
TYPE ST_EL1918 :
STRUCT
	//--------------------------------------------------------------------------------------------------------
	sTerminalName                                           :   STRING(200):= 'EL1918 | 8-Channel Safety Digital Input';
    //============================================================================================================================	
	// TERMINAL - EL1918 8-Channel Digital Input Terminal (Term 4)	
	iEL1918_Ch1                			AT %I*			: 	BOOL;	// EL1918 channel 1
	iEL1918_Ch2                   		AT %I*			: 	BOOL;	// EL1918 channel 2
	iEL1918_Ch3        					AT %I*	 		: 	BOOL;	// EL1918 channel 3
	iEL1918_Ch4   						AT %I*	 		: 	BOOL;	// EL1918 channel 4
	iEL1918_Ch5         				AT %I*	 		: 	BOOL;	// EL1918 channel 5 		     			
	iEL1918_Ch6 						AT %I*			: 	BOOL;	// EL1918 channel 6
	iEL1918_Ch7               			AT %I*          :   BOOL;   // EL1918 channel 7 
    iEL1918_Ch8          				AT %I*          :   BOOL;   // EL1918 channel 8
 		
	stTerminalInfo											: 	ST_Terminal_Info;

END_STRUCT
END_TYPE

// ---- DUTs/04_IO_Mapping/Terminals/ST_EL2502.TcDUT
TYPE ST_EL2502 :
STRUCT
	sTerminalName : STRING(80) := 'EL2502 | 2-Channel PWM Output';

    iEL2502_Ch1  AT %Q* : UINT;
    iEL2502_Ch2  AT %Q* : UINT;

    stTerminalInfo : ST_Terminal_Info;
END_STRUCT
END_TYPE

// ---- DUTs/04_IO_Mapping/Terminals/ST_EL2904.TcDUT
TYPE ST_EL2904 :
STRUCT
    sTerminalName : STRING(80) := 'EL2904 | 4-Channel TwinSAFE Digital Output';

    // Diagnostic representation only. Functional commands are exchanged
    // through GVL_Safety aliases and evaluated inside the TwinSAFE project.
    bOutput : ARRAY[1..4] OF BOOL;
    bError  : BOOL;
    bReady  : BOOL;

    stTerminalInfo : ST_Terminal_Info;
END_STRUCT
END_TYPE

// ---- DUTs/04_IO_Mapping/Terminals/ST_EL3058.TcDUT
TYPE ST_EL3058 :
STRUCT
	//--------------------------------------------------------------------------------------------------------
	sTerminalName                                           :   STRING(200):= 'EL3058 | 8-Channel Analog Input 4..20mA';
    //============================================================================================================================	
	// TERMINAL - EL3058 4-Channel Analog Input Terminal (Term 11)	
	iEL3058_Ch1               				AT %I*			: 	UINT;	// EL1809 channel 1
	iEL3058_Ch2                   			AT %I*			: 	UINT;	// EL1809 channel 2
	iEL3058_Ch3        						AT %I*	 		: 	UINT;	// EL1809 channel 3
	iEL3058_Ch4	   							AT %I*	 		: 	UINT;	// EL1809 channel 4
	iEL3058_Ch5	   							AT %I*	 		: 	UINT;	// EL1809 channel 5
	iEL3058_Ch6	   							AT %I*	 		: 	UINT;	// EL1809 channel 6
	iEL3058_Ch7	   							AT %I*	 		: 	UINT;	// EL1809 channel 7
	iEL3058_Ch8	   							AT %I*	 		: 	UINT;	// EL1809 channel 8
	
	stTerminalInfo											: 	ST_Terminal_Info;

END_STRUCT
END_TYPE

// ---- DUTs/04_IO_Mapping/Terminals/ST_EL3064.TcDUT
TYPE ST_EL3064 :
STRUCT
	//--------------------------------------------------------------------------------------------------------
	sTerminalName                                           :   STRING(200):= 'EL3064 | 4-Channel Analog Input 0..10V';
    //============================================================================================================================	
	// TERMINAL - EL3058 4-Channel Analog Input Terminal (Term 11)	
	iEL3064_Ch1               				AT %I*			: 	UINT;	// EL1809 channel 1
	iEL3064_Ch2                   			AT %I*			: 	UINT;	// EL1809 channel 2
	iEL3064_Ch3        						AT %I*	 		: 	UINT;	// EL1809 channel 3
	iEL3064_Ch4	   							AT %I*	 		: 	UINT;	// EL1809 channel 4
	
	stTerminalInfo											: 	ST_Terminal_Info;

END_STRUCT
END_TYPE

// ---- DUTs/04_IO_Mapping/Terminals/ST_EL6910.TcDUT
TYPE ST_EL6910 :
STRUCT
	
	// TERMINAL - EL6910	TwinSAFE logic	 (Term 3)
	sTerminalName                                           :   STRING(200):= 'EL6910 | TwinSAFE logic';
	stTerminalInfo											: 	ST_Terminal_Info;

END_STRUCT
END_TYPE

// ---- DUTs/04_IO_Mapping/Terminals/ST_EL7201.TcDUT
TYPE ST_EL7201 :
STRUCT
	sTerminalName : STRING(80) := 'EL7201-9014 | 1-Channel Servomotor - Axis 1 [Reel Payout]';

    stTerminalInfo : ST_Terminal_Info;
END_STRUCT
END_TYPE

// ---- DUTs/05_AlarmsAndEvents/E_AlarmId.TcDUT
{attribute 'qualified_only'}
{attribute 'strict'}
{attribute 'to_string'}
TYPE E_AlarmId :
(
    None := 0,
    SafetyNotAvailable := 1000,
    EmergencyStopActive := 1001,
    MainDoorNotSafe := 1002,
    LeftFlapSafetyActive := 1003,
    RightFlapSafetyActive := 1004,
    FsoeNotHealthy := 1005,
    SafetyLogicNotHealthy := 1006,
    IndexFault := 2000,
    IndexPositionInvalid := 2001,
    IndexWrongPositionTimeout := 2002,
    ProcessCylinderFault := 3000,
    ProcessEquipmentFault := 3001,
    PuckRemovedWhileLocked := 4000,
    PuckSensorMismatch := 4001,
    OperatorExchangeFault := 5000,
    RejectConfirmationRequired := 5001,
    ProcessedPartRemovalRequired := 5002,
    InitialisationTimeout := 6000,
    StoppingTimeout := 6001
);
END_TYPE

// ---- DUTs/05_AlarmsAndEvents/E_AlarmSeverity.TcDUT
{attribute 'qualified_only'}
{attribute 'strict'}
{attribute 'to_string'}
TYPE E_AlarmSeverity :
(
    Information := 0,
    Warning := 10,
    Fault := 20,
    SafetyStop := 30
);
END_TYPE

// ---- DUTs/05_AlarmsAndEvents/E_MachineAlarm.TcDUT
{attribute 'qualified_only'}
{attribute 'strict'}
TYPE E_MachineAlarm :
(
    None := 0,
    EmergencyStop := 1000,
    MainDoorSafety := 1001,
    LeftSafetyFlap := 1002,
    RightSafetyFlap := 1003,
    Up24VSupply := 1100,
    Us24VSupply := 1101,
    Up48VSupply := 1102,
    AirSupply := 1200,
    IndexFault := 1300,
    InitialisationTimeout := 1400,
    StoppingTimeout := 1401
);
END_TYPE

// ---- DUTs/05_AlarmsAndEvents/ST_ActiveEvents.TcDUT
TYPE ST_ActiveEvents :
STRUCT
	
	sEventTex									: STRING(255);
	sType										: STRING(255);
	sSolution									: STRING(255);
	abType										: DINT;					//1:Alarm
																		//2:Alert
																		//3:Message
END_STRUCT
END_TYPE

// ---- DUTs/05_AlarmsAndEvents/ST_AlarmManagerStatus.TcDUT
TYPE ST_AlarmManagerStatus :
STRUCT
    bHasFault             : BOOL;
    bHasSafetyStopFault   : BOOL;
    uiActiveCount         : UINT;
    eHighestAlarm         : E_AlarmId;
    aActive               : ARRAY[1..20] OF ST_ActiveAlarm;
END_STRUCT
END_TYPE

// ---- DUTs/05_AlarmsAndEvents/ST_EVENT.TcDUT
TYPE ST_EVENT :
STRUCT
	bFault								: BOOL;
	bCycleStopRequest					: BOOL;
	bMessage							: BOOL;
	bPersistentMessage				: BOOL; // Live message; clears only when condition becomes FALSE
	
	bAssignedID							: DINT;
	
	bEventFlag							: BOOL;
	bEventTimer							: TON;
	bEventText							: STRING(255);
	bEventTextHMI						: STRING(255);
	sSolution							: STRING(255);
	bActive								: BOOL;
END_STRUCT
END_TYPE

// ---- DUTs/05_AlarmsAndEvents/ST_EventsAssigment.TcDUT
TYPE ST_EventsAssigment :
STRUCT
	sEventText	: STRING(255);
	sSolution	: STRING(255);
END_STRUCT
END_TYPE

// ---- DUTs/05_AlarmsAndEvents/ST_StationEvents.TcDUT
TYPE ST_StationEvents :
STRUCT
	aEvents								: ARRAY [0..100] OF ST_EVENT;	
	
	bFault								: BOOL;
	bCycleStopRequest					: BOOL;
END_STRUCT
END_TYPE

// ---- GVLs/GVL_Config.TcGVL
{attribute 'qualified_only'}
VAR_GLOBAL PERSISTENT RETAIN
    stMachine : ST_MachineConfig := (
        tInitialiseTimeout := T#20S,
        tStoppingTimeout := T#15S,
        tIndexTimeout := T#10S,
        eOperatorPosition := E_TablePosition.Position1,
        ePatchDispensePosition := E_TablePosition.Position2,
        eHeatStakePosition := E_TablePosition.Position3,
        eVisionPosition := E_TablePosition.Position4,
        eRejectPosition := E_TablePosition.Position1,
        bAllowEmptyNestIndex := TRUE,
        bRequireRejectConfirm := TRUE
    );
    aNestEnabled : ARRAY[1..4] OF BOOL := [TRUE, TRUE, TRUE, TRUE];
END_VAR

// ---- GVLs/GVL_EtherCAT.TcGVL
{attribute 'qualified_only'}
VAR_GLOBAL
    stTerm1_EK1100   : ST_EK1100;
    stTerm2_EL6070   : ST_EL6070;
    stTerm3_EL6910   : ST_EL6910;
    stTerm4_EL1918   : ST_EL1918;
    stTerm5_EL1918   : ST_EL1918;
    stTerm6_EL2904   : ST_EL2904;
    stTerm7_EL1809   : ST_EL1809;
    stTerm8_EL1809   : ST_EL1809;
    stTerm9_EL2809   : ST_EL2809;
    stTerm10_EL2809  : ST_EL2809;
    stTerm11_EL3058  : ST_EL3058;
	stTerm13_EL2502  : ST_EL2502;
	stTerm15_EL7201  : ST_EL7201;
	stTerm16_EL7201  : ST_EL7201;
	stTerm17_EL7201  : ST_EL7201;
	stTerm18_EL2904  : ST_EL2904;
    stTerm19_EL1809  : ST_EL1809;
	stTerm20_EL3314  : ST_EL3314;
	stTerm21_EL6633  : ST_EL6633;
END_VAR

// ---- GVLs/GVL_HMI.TcGVL
{attribute 'qualified_only'}
VAR_GLOBAL
    stCommands : ST_HmiCommands;
    stStatus : ST_HmiStatus;
    StatusHMI : ST_StatusBanner;
    astActiveEvents : ARRAY[0..50] OF ST_ActiveEvents;
    astEventsHistory : ARRAY[0..200] OF ST_EventsHistory;
    astTestHistory : ARRAY[0..2000] OF ST_TestHistory;
    stEventsAssigment : ST_EventsAssigmentGeneral;
    sSystemTime : STRING(255);
    sSystemDate : STRING(255);
    stStatistics : ST_HmiStatistics;
    bBlink_1Hz : BOOL;
    bHMIAlive : BOOL;
END_VAR
VAR_GLOBAL CONSTANT
    sWHITE : STRING(40) := '{"color":"rgba(255,255,255,255)"}';
    sBLACK : STRING(40) := '{"color":"rgba(0,0,0,1)"}';
    sYELLOW : STRING(40) := '{"color":"rgba(255,255,0,1)"}';
    sGREEN : STRING(40) := '{"color":"rgba(70,166,63,1)"}';
    sRED : STRING(40) := '{"color":"rgba(255,0,0,1)"}';
    sBLUEInProgress : STRING(40) := '{"color":"rgba(54,100,221,1)"}';
    sGREY : STRING(40) := '{"color":"rgba(164,158,158,1)"}';
    sDARKGREY : STRING(40) := '{"color":"rgba(50,50,50,1)"}';
    sTRANSP : STRING(40) := '{"color":"rgba(255,255,255,0)"}';
    sREDFail : STRING(40) := '{"color":"rgba(244,68,68,255)"}';
    sSystemName : STRING := 'Patch Press';
    sApplication : STRING := 'Patch Press Machine';
    sProjectID : STRING := 'TE1108';
    sSoftwareVersion : STRING := 'v0.1.0-foundation';
END_VAR

// ---- GVLs/GVL_MASTER.TcGVL
{attribute 'qualified_only'}
VAR_GLOBAL
    stInputs  : ST_MachineInputs;
    stOutputs : ST_MachineOutputs;
    stCommand : ST_MachineCommand;
    stStatus  : ST_MachineStatus;
    stStationEvents   : ARRAY[0..4] OF ST_StationEvents;
    stEventsAssigment : ST_EventsAssigmentGeneral;
    astActiveEvents   : ARRAY[0..50] OF ST_ActiveEvents;
    sSystemTime       : STRING(255);
    sSystemDate       : STRING(255);
    bMachineFault     : BOOL;
    bCycleStopRequest : BOOL;
END_VAR

// ---- GVLs/GVL_Motion.TcGVL
{attribute 'qualified_only'}
VAR_GLOBAL
    // Term 15 - EL7201-9014 - Axis 1 - Reel Payout
    AxisReelPayout      : ST_Axis;

    // Term 16 - EL7201-9014 - Axis 2 - Material Index
    AxisMaterialIndex   : ST_Axis;

    // Term 17 - EL7201-9014 - Axis 3 - Slack
    AxisSlack           : ST_Axis;
END_VAR

// ---- GVLs/GVL_PatchPress_Interface.TcGVL
{attribute 'qualified_only'}
VAR_GLOBAL
    bPatchDispenseCommissioned : BOOL := FALSE;
    bHeatStakeCommissioned     : BOOL := FALSE;
    bVisionCommissioned        : BOOL := FALSE;
    // Engineering-only mode for commissioning the validated core before the
    // three process stations are available. Keep FALSE for production.
    bCoreCommissioningMode     : BOOL := FALSE;
END_VAR

// ---- GVLs/GVL_Persistent.TcGVL
{attribute 'qualified_only'}
VAR_GLOBAL PERSISTENT RETAIN
    astEventsHistory : ARRAY[0..200] OF ST_EventsHistory;
END_VAR

// ---- GVLs/GVL_Safety.TcGVL
{attribute 'qualified_only'}
VAR_GLOBAL
    // ---------------------------------------------------------------------
    // TwinSAFE -> standard PLC aliases (link as PLC inputs in the Safety
    // project). These are validated statuses/diagnostics, not reconstructed
    // safety logic in the standard PLC.
    // ---------------------------------------------------------------------
    bSafetyOk                  AT %I* : BOOL;
    bEmergencyStopOk           AT %I* : BOOL;
    bMainDoorUnSafe            AT %I* : BOOL;
    bLeftFlapSafe              AT %I* : BOOL;
    bRightFlapSafe             AT %I* : BOOL;
    bFlapsSafe                 AT %I* : BOOL;
    bTwoHandSafe               AT %I* : BOOL;
    bAirSupplySafe             AT %I* : BOOL;
    bFsoeOk                    AT %I* : BOOL;
    bSafetyLogicOk             AT %I* : BOOL;

    // Diagnostic/command feedback exported by TwinSAFE.
    bResetButtonPressed        AT %I* : BOOL;
    bMainDoorClosed            AT %I* : BOOL;
    bMainDoorLocked            AT %I* : BOOL;
    bMainDoorDiagnosticOk      AT %I* : BOOL;
    bMs6FeedbackOk             AT %I* : BOOL;
    bAirExhausted              AT %I* : BOOL;

    // ---------------------------------------------------------------------
    // Standard PLC -> TwinSAFE request aliases (link as PLC outputs in the
    // Safety project). TwinSAFE remains the owner of EL2904 safe outputs.
    // ---------------------------------------------------------------------
    bSafetyRunRequest          AT %Q* : BOOL;
    bSafetyResetRequest        AT %Q* : BOOL;
    bAirSupplyEnableRequest    AT %Q* : BOOL;
    bMainDoorLockRequest       AT %Q* : BOOL;
	bMachineFaultRequest 			  : BOOL;
	bSafetyErrorAcknowledgementRequest : BOOL;
	
	
END_VAR

// ---- POUs/MAIN.TcPOU
PROGRAM MAIN
VAR
END_VAR

PRG_TerminalMapping.ReadInputs();
PRG_ReadInputs();
PRG_HmiCommands();
PRG_Main();
PRG_Events();
PRG_HmiStatus();
PRG_WriteOutputs();
PRG_TerminalMapping.WriteOutputs();

END_PROGRAM

// ---- POUs/04_IO_Mapping/PRG_TerminalMapping.TcPOU
PROGRAM PRG_TerminalMapping
VAR
    uiIndexPositionCode : UINT;
END_VAR

METHOD PUBLIC ReadInputs
GVL_IO.stInputs.bEmergencyStopChannel1 := GVL_EtherCAT.stTerm4_EL1918.iEL1918_Ch1;
GVL_IO.stInputs.bEmergencyStopChannel2 := GVL_EtherCAT.stTerm4_EL1918.iEL1918_Ch2;
GVL_IO.stInputs.bResetButton := GVL_EtherCAT.stTerm4_EL1918.iEL1918_Ch3;
GVL_IO.stInputs.bMainDoorChannel1 := GVL_EtherCAT.stTerm4_EL1918.iEL1918_Ch4;
GVL_IO.stInputs.bMainDoorChannel2 := GVL_EtherCAT.stTerm4_EL1918.iEL1918_Ch5;
GVL_IO.stInputs.bMainDoorFeedback := GVL_EtherCAT.stTerm4_EL1918.iEL1918_Ch6;
GVL_IO.stInputs.bMs6FeedbackOk := GVL_EtherCAT.stTerm4_EL1918.iEL1918_Ch7;
GVL_IO.stInputs.bAirExhausted := GVL_EtherCAT.stTerm4_EL1918.iEL1918_Ch8;
GVL_IO.stInputs.bTouchButtonLeft := GVL_EtherCAT.stTerm5_EL1918.iEL1918_Ch3;
GVL_IO.stInputs.bTouchButtonRight := GVL_EtherCAT.stTerm5_EL1918.iEL1918_Ch4;
GVL_IO.stInputs.bRightFlapChannel1 := GVL_EtherCAT.stTerm5_EL1918.iEL1918_Ch5;
GVL_IO.stInputs.bRightFlapChannel2 := GVL_EtherCAT.stTerm5_EL1918.iEL1918_Ch6;
GVL_IO.stInputs.bLeftFlapChannel1 := GVL_EtherCAT.stTerm5_EL1918.iEL1918_Ch7;
GVL_IO.stInputs.bLeftFlapChannel2 := GVL_EtherCAT.stTerm5_EL1918.iEL1918_Ch8;
GVL_IO.stInputs.bStartButton := GVL_EtherCAT.stTerm7_EL1809.iEL1809_Ch1;
GVL_IO.stInputs.bStopButton := NOT GVL_EtherCAT.stTerm7_EL1809.iEL1809_Ch2;
GVL_IO.stInputs.bUp24VPowerSupplyOk := GVL_EtherCAT.stTerm7_EL1809.iEL1809_Ch3;
GVL_IO.stInputs.bUs24VPowerSupplyOk := GVL_EtherCAT.stTerm7_EL1809.iEL1809_Ch4;
GVL_IO.stInputs.b48VPowerSupplyOk := GVL_EtherCAT.stTerm7_EL1809.iEL1809_Ch5;
GVL_IO.stInputs.bIndexPositionSensor1 := GVL_EtherCAT.stTerm7_EL1809.iEL1809_Ch6;
GVL_IO.stInputs.bIndexPositionSensor2 := GVL_EtherCAT.stTerm7_EL1809.iEL1809_Ch7;
GVL_IO.stInputs.bIndexPositionSensor3 := GVL_EtherCAT.stTerm7_EL1809.iEL1809_Ch8;
GVL_IO.stInputs.bIndexCompletedSensor := GVL_EtherCAT.stTerm7_EL1809.iEL1809_Ch9;
GVL_IO.stInputs.bIndexLocked := GVL_EtherCAT.stTerm7_EL1809.iEL1809_Ch10;
GVL_IO.stInputs.bIndexReady := GVL_EtherCAT.stTerm7_EL1809.iEL1809_Ch11;
GVL_IO.stInputs.bLoadingStationEaglePresent := GVL_EtherCAT.stTerm7_EL1809.iEL1809_Ch12;
GVL_IO.stInputs.bRejectChutePartPresent := GVL_EtherCAT.stTerm7_EL1809.iEL1809_Ch13;
GVL_IO.stInputs.bHeatStakeEaglePresent := GVL_EtherCAT.stTerm7_EL1809.iEL1809_Ch14;
GVL_IO.stInputs.bHeatStakePatchPresent := GVL_EtherCAT.stTerm7_EL1809.iEL1809_Ch15;
GVL_IO.stInputs.bPbupMagnetPresent := GVL_EtherCAT.stTerm7_EL1809.iEL1809_Ch16;
uiIndexPositionCode := 0;
IF GVL_IO.stInputs.bIndexPositionSensor1 THEN uiIndexPositionCode := uiIndexPositionCode + 1; END_IF
IF GVL_IO.stInputs.bIndexPositionSensor2 THEN uiIndexPositionCode := uiIndexPositionCode + 2; END_IF
IF GVL_IO.stInputs.bIndexPositionSensor3 THEN uiIndexPositionCode := uiIndexPositionCode + 4; END_IF
IF GVL_IO.stInputs.bIndexLocked THEN GVL_IO.stInputs.eIndexPosition := UINT_TO_E_TablePosition(uiIndexPositionCode); ELSE GVL_IO.stInputs.eIndexPosition := E_TablePosition.Unknown; END_IF
GVL_IO.stInputs.bStation1SupportRetracted := GVL_EtherCAT.stTerm8_EL1809.iEL1809_Ch1;
GVL_IO.stInputs.bStation1SupportExtended := GVL_EtherCAT.stTerm8_EL1809.iEL1809_Ch2;
GVL_IO.stInputs.bStation2SupportRetracted := GVL_EtherCAT.stTerm8_EL1809.iEL1809_Ch3;
GVL_IO.stInputs.bStation2SupportExtended := GVL_EtherCAT.stTerm8_EL1809.iEL1809_Ch4;
GVL_IO.stInputs.bStation3SupportRetracted := GVL_EtherCAT.stTerm8_EL1809.iEL1809_Ch5;
GVL_IO.stInputs.bStation3SupportExtended := GVL_EtherCAT.stTerm8_EL1809.iEL1809_Ch6;
GVL_IO.stInputs.bHorizontalMiniSlideRetracted := GVL_EtherCAT.stTerm8_EL1809.iEL1809_Ch7;
GVL_IO.stInputs.bHorizontalMiniSlideExtended := GVL_EtherCAT.stTerm8_EL1809.iEL1809_Ch8;
GVL_IO.stInputs.bVerticalMiniSlideRetracted := GVL_EtherCAT.stTerm8_EL1809.iEL1809_Ch9;
GVL_IO.stInputs.bVerticalMiniSlideExtended := GVL_EtherCAT.stTerm8_EL1809.iEL1809_Ch10;
GVL_IO.stInputs.bIntermediateModuleRetracted := GVL_EtherCAT.stTerm8_EL1809.iEL1809_Ch11;
GVL_IO.stInputs.bIntermediateModuleExtended := GVL_EtherCAT.stTerm8_EL1809.iEL1809_Ch12;
GVL_IO.stInputs.bRotaryGripperOpened := GVL_EtherCAT.stTerm8_EL1809.iEL1809_Ch13;
GVL_IO.stInputs.bRotaryGripperClosed := GVL_EtherCAT.stTerm8_EL1809.iEL1809_Ch14;
GVL_IO.stInputs.bRotaryGripperPick0 := GVL_EtherCAT.stTerm8_EL1809.iEL1809_Ch15;
GVL_IO.stInputs.bRotaryGripperPlace180 := GVL_EtherCAT.stTerm8_EL1809.iEL1809_Ch16;
GVL_IO.stInputs.bMembraneTransferRetracted := GVL_EtherCAT.stTerm19_EL1809.iEL1809_Ch9;
GVL_IO.stInputs.bMembraneTransferExtended := GVL_EtherCAT.stTerm19_EL1809.iEL1809_Ch10;
GVL_IO.stInputs.bMiddleRockerDown := GVL_EtherCAT.stTerm19_EL1809.iEL1809_Ch11;
GVL_IO.stInputs.bMiddleRockerUp := GVL_EtherCAT.stTerm19_EL1809.iEL1809_Ch12;
GVL_IO.stInputs.bBottomRockerDown := GVL_EtherCAT.stTerm19_EL1809.iEL1809_Ch13;
GVL_IO.stInputs.bBottomRockerUp := GVL_EtherCAT.stTerm19_EL1809.iEL1809_Ch14;
GVL_IO.stInputs.bTopRockerDown := GVL_EtherCAT.stTerm19_EL1809.iEL1809_Ch15;
GVL_IO.stInputs.bTopRockerUp := GVL_EtherCAT.stTerm19_EL1809.iEL1809_Ch16;
GVL_IO.stInputs.uiMainAirPressureRaw := GVL_EtherCAT.stTerm11_EL3058.iEL3058_Ch1;
GVL_IO.stInputs.uiPressureRegulatorActualRaw := GVL_EtherCAT.stTerm11_EL3058.iEL3058_Ch2;
GVL_IO.stInputs.bSafetyOk := GVL_Safety.bSafetyOk;
GVL_IO.stInputs.bTwoHandsSafe := GVL_Safety.bTwoHandSafe;
GVL_IO.stInputs.bMainDoorClosed := GVL_Safety.bMainDoorClosed;
GVL_IO.stInputs.bMainDoorLocked := GVL_Safety.bMainDoorLocked;
GVL_IO.stInputs.bMainDoorUnsafe := GVL_Safety.bMainDoorUnSafe;
GVL_IO.stInputs.bMainDoorDiagnosticOk := GVL_Safety.bMainDoorDiagnosticOk;
END_METHOD

METHOD PUBLIC WriteOutputs
GVL_Safety.bSafetyRunRequest := GVL_IO.stOutputs.bSafetyRunRequest;
GVL_Safety.bSafetyResetRequest := GVL_IO.stOutputs.bSafetyResetRequest;
GVL_Safety.bSafetyErrorAcknowledgementRequest := GVL_IO.stOutputs.bSafetyErrorAcknowledgementRequest;
GVL_Safety.bAirSupplyEnableRequest := GVL_IO.stOutputs.bAirSupplyEnable;
GVL_Safety.bMainDoorLockRequest := GVL_IO.stOutputs.bMainDoorLockRequest;
GVL_EtherCAT.stTerm9_EL2809.iEL2809_Ch1 := GVL_IO.stOutputs.bLedStart;
GVL_EtherCAT.stTerm9_EL2809.iEL2809_Ch2 := GVL_IO.stOutputs.bLedReset;
GVL_EtherCAT.stTerm9_EL2809.iEL2809_Ch3 := GVL_IO.stOutputs.bStatusIndicator;
GVL_EtherCAT.stTerm9_EL2809.iEL2809_Ch4 := GVL_IO.stOutputs.bInternalLight;
GVL_EtherCAT.stTerm9_EL2809.iEL2809_Ch5 := GVL_IO.stOutputs.bNestLight;

// Temporary assumption for Patch Press commissioning:
// Reuse the validated Silicone Station index valve mapping on Term 10.
GVL_EtherCAT.stTerm10_EL2809.iEL2809_Ch1 := GVL_IO.stOutputs.bIndexStopPortB;
GVL_EtherCAT.stTerm10_EL2809.iEL2809_Ch2 := GVL_IO.stOutputs.bIndexRotatePortA;
END_METHOD

END_PROGRAM

// ---- POUs/02_Components/Index/UINT_TO_E_TablePosition.TcPOU
FUNCTION UINT_TO_E_TablePosition : E_TablePosition
VAR_INPUT
    uiPosition : UINT;
END_VAR

CASE uiPosition OF
    1:
        UINT_TO_E_TablePosition := E_TablePosition.Position1;

    2:
        UINT_TO_E_TablePosition := E_TablePosition.Position2;

    3:
        UINT_TO_E_TablePosition := E_TablePosition.Position3;

    4:
        UINT_TO_E_TablePosition := E_TablePosition.Position4;

ELSE
    UINT_TO_E_TablePosition := E_TablePosition.Unknown;
END_CASE

END_FUNCTION

// ---- POUs/00_Application/PRG_ReadInputs.TcPOU
PROGRAM PRG_ReadInputs
VAR
END_VAR

GVL_MASTER.stInputs.bStartButton := GVL_IO.stInputs.bStartButton;
GVL_MASTER.stInputs.bStopButton := GVL_IO.stInputs.bStopButton;
GVL_MASTER.stInputs.bResetButton := GVL_IO.stInputs.bResetButton;
GVL_MASTER.stInputs.bTwoHandsSafe := GVL_IO.stInputs.bTwoHandsSafe;
GVL_MASTER.stInputs.bTouchButtonLeft := GVL_IO.stInputs.bTouchButtonLeft;
GVL_MASTER.stInputs.bTouchButtonRight := GVL_IO.stInputs.bTouchButtonRight;
GVL_MASTER.stInputs.bUp24VPowerSupplyOk := GVL_IO.stInputs.bUp24VPowerSupplyOk;
GVL_MASTER.stInputs.bUs24VPowerSupplyOk := GVL_IO.stInputs.bUs24VPowerSupplyOk;
GVL_MASTER.stInputs.b48VPowerSupplyOk := GVL_IO.stInputs.b48VPowerSupplyOk;
GVL_MASTER.stInputs.bEmergencyStopChannel1 := GVL_IO.stInputs.bEmergencyStopChannel1;
GVL_MASTER.stInputs.bEmergencyStopChannel2 := GVL_IO.stInputs.bEmergencyStopChannel2;
GVL_MASTER.stInputs.bMainDoorChannel1 := GVL_IO.stInputs.bMainDoorChannel1;
GVL_MASTER.stInputs.bMainDoorChannel2 := GVL_IO.stInputs.bMainDoorChannel2;
GVL_MASTER.stInputs.bMainDoorFeedback := GVL_IO.stInputs.bMainDoorFeedback;
GVL_MASTER.stInputs.bLeftFlapChannel1 := GVL_IO.stInputs.bLeftFlapChannel1;
GVL_MASTER.stInputs.bLeftFlapChannel2 := GVL_IO.stInputs.bLeftFlapChannel2;
GVL_MASTER.stInputs.bRightFlapChannel1 := GVL_IO.stInputs.bRightFlapChannel1;
GVL_MASTER.stInputs.bRightFlapChannel2 := GVL_IO.stInputs.bRightFlapChannel2;
GVL_MASTER.stInputs.bMainDoorClosed := GVL_IO.stInputs.bMainDoorClosed;
GVL_MASTER.stInputs.bMainDoorLocked := GVL_IO.stInputs.bMainDoorLocked;
GVL_MASTER.stInputs.bMainDoorUnsafe := GVL_IO.stInputs.bMainDoorUnsafe;
GVL_MASTER.stInputs.bMainDoorDiagnosticOk := GVL_IO.stInputs.bMainDoorDiagnosticOk;
GVL_MASTER.stInputs.bMs6FeedbackOk := GVL_IO.stInputs.bMs6FeedbackOk;
GVL_MASTER.stInputs.bAirExhausted := GVL_IO.stInputs.bAirExhausted;
GVL_MASTER.stInputs.stSafety.bSafetyOk := GVL_IO.stInputs.bSafetyOk;
GVL_MASTER.stInputs.stSafety.bMotionSafetyPermitted := GVL_IO.stInputs.bSafetyOk;
GVL_MASTER.stInputs.stSafety.bProcessSafetyPermitted := GVL_IO.stInputs.bSafetyOk;
GVL_MASTER.stInputs.stSafety.bMainDoorSafe := NOT GVL_IO.stInputs.bMainDoorUnsafe;
GVL_MASTER.stInputs.stSafety.bLeftFlapSafe := GVL_Safety.bLeftFlapSafe;
GVL_MASTER.stInputs.stSafety.bRightFlapSafe := GVL_Safety.bRightFlapSafe;
GVL_MASTER.stInputs.bEventFault := GVL_MASTER.bMachineFault;
GVL_MASTER.stInputs.bEventCycleStopRequest := GVL_MASTER.bCycleStopRequest;
GVL_MASTER.stInputs.bIndexReady := GVL_IO.stInputs.bIndexReady;
GVL_MASTER.stInputs.bIndexLocked := GVL_IO.stInputs.bIndexLocked;
GVL_MASTER.stInputs.bIndexCompletedSensor := GVL_IO.stInputs.bIndexCompletedSensor;
GVL_MASTER.stInputs.eIndexPosition := GVL_IO.stInputs.eIndexPosition;
GVL_MASTER.stInputs.bLoadingStationEaglePresent := GVL_IO.stInputs.bLoadingStationEaglePresent;
GVL_MASTER.stInputs.bRejectChutePartPresent := GVL_IO.stInputs.bRejectChutePartPresent;
GVL_MASTER.stInputs.bHeatStakeEaglePresent := GVL_IO.stInputs.bHeatStakeEaglePresent;
GVL_MASTER.stInputs.bHeatStakePatchPresent := GVL_IO.stInputs.bHeatStakePatchPresent;
GVL_MASTER.stInputs.bPbupMagnetPresent := GVL_IO.stInputs.bPbupMagnetPresent;
GVL_MASTER.stInputs.bStation1SupportRetracted := GVL_IO.stInputs.bStation1SupportRetracted;
GVL_MASTER.stInputs.bStation1SupportExtended := GVL_IO.stInputs.bStation1SupportExtended;
GVL_MASTER.stInputs.bStation2SupportRetracted := GVL_IO.stInputs.bStation2SupportRetracted;
GVL_MASTER.stInputs.bStation2SupportExtended := GVL_IO.stInputs.bStation2SupportExtended;
GVL_MASTER.stInputs.bStation3SupportRetracted := GVL_IO.stInputs.bStation3SupportRetracted;
GVL_MASTER.stInputs.bStation3SupportExtended := GVL_IO.stInputs.bStation3SupportExtended;
GVL_MASTER.stInputs.bHorizontalMiniSlideRetracted := GVL_IO.stInputs.bHorizontalMiniSlideRetracted;
GVL_MASTER.stInputs.bHorizontalMiniSlideExtended := GVL_IO.stInputs.bHorizontalMiniSlideExtended;
GVL_MASTER.stInputs.bVerticalMiniSlideRetracted := GVL_IO.stInputs.bVerticalMiniSlideRetracted;
GVL_MASTER.stInputs.bVerticalMiniSlideExtended := GVL_IO.stInputs.bVerticalMiniSlideExtended;
GVL_MASTER.stInputs.bIntermediateModuleRetracted := GVL_IO.stInputs.bIntermediateModuleRetracted;
GVL_MASTER.stInputs.bIntermediateModuleExtended := GVL_IO.stInputs.bIntermediateModuleExtended;
GVL_MASTER.stInputs.bRotaryGripperOpened := GVL_IO.stInputs.bRotaryGripperOpened;
GVL_MASTER.stInputs.bRotaryGripperClosed := GVL_IO.stInputs.bRotaryGripperClosed;
GVL_MASTER.stInputs.bRotaryGripperPick0 := GVL_IO.stInputs.bRotaryGripperPick0;
GVL_MASTER.stInputs.bRotaryGripperPlace180 := GVL_IO.stInputs.bRotaryGripperPlace180;
GVL_MASTER.stInputs.bMembraneTransferRetracted := GVL_IO.stInputs.bMembraneTransferRetracted;
GVL_MASTER.stInputs.bMembraneTransferExtended := GVL_IO.stInputs.bMembraneTransferExtended;
GVL_MASTER.stInputs.bMiddleRockerDown := GVL_IO.stInputs.bMiddleRockerDown;
GVL_MASTER.stInputs.bMiddleRockerUp := GVL_IO.stInputs.bMiddleRockerUp;
GVL_MASTER.stInputs.bBottomRockerDown := GVL_IO.stInputs.bBottomRockerDown;
GVL_MASTER.stInputs.bBottomRockerUp := GVL_IO.stInputs.bBottomRockerUp;
GVL_MASTER.stInputs.bTopRockerDown := GVL_IO.stInputs.bTopRockerDown;
GVL_MASTER.stInputs.bTopRockerUp := GVL_IO.stInputs.bTopRockerUp;
GVL_MASTER.stInputs.uiMainAirPressureRaw := GVL_IO.stInputs.uiMainAirPressureRaw;
GVL_MASTER.stInputs.uiPressureRegulatorActualRaw := GVL_IO.stInputs.uiPressureRegulatorActualRaw;

END_PROGRAM

// ---- POUs/00_Application/PRG_HmiCommands.TcPOU
PROGRAM PRG_HmiCommands
VAR
    rtStart : R_TRIG;
    rtReset : R_TRIG;
    rtAck : R_TRIG;
END_VAR

rtStart(CLK := GVL_MASTER.stInputs.bStartButton OR GVL_HMI.stCommands.bStart);
rtReset(CLK := GVL_MASTER.stInputs.bResetButton OR GVL_HMI.stCommands.bReset);
rtAck(CLK := GVL_HMI.stCommands.bAcknowledge);
GVL_MASTER.stCommand.bStart := rtStart.Q;
GVL_MASTER.stCommand.bStop := GVL_MASTER.stInputs.bStopButton OR GVL_HMI.stCommands.bStop;
GVL_MASTER.stCommand.bReset := rtReset.Q;
GVL_MASTER.stCommand.bAcknowledge := rtAck.Q;
GVL_MASTER.stCommand.bManualRequest := GVL_HMI.stCommands.bManualRequest;
GVL_MASTER.stCommand.bIndexerManualEnable := GVL_HMI.stCommands.bIndexerManualEnable;
GVL_MASTER.stCommand.bManualIndexForward := GVL_HMI.stCommands.bManualIndexForward;
GVL_MASTER.stCommand.bManualIndexHome := GVL_HMI.stCommands.bManualIndexHome;
GVL_MASTER.stCommand.bManualMainDoorUnlock := GVL_HMI.stCommands.bManualMainDoorUnlock;
GVL_MASTER.stCommand.uiResetStatisticsNestId := GVL_HMI.stCommands.uiResetStatisticsNestId;

END_PROGRAM

// ---- POUs/00_Application/PRG_Main.TcPOU
PROGRAM PRG_Main
VAR
    fbMachine : FB_IndexedPatchPressMachine;
END_VAR

fbMachine.Cyclic(
    stInputs := GVL_MASTER.stInputs,
    stCommand := GVL_MASTER.stCommand,
    stConfig := GVL_Config.stMachine,
    bPatchDispenseCommissioned := GVL_PatchPress_Interface.bPatchDispenseCommissioned,
    bHeatStakeCommissioned := GVL_PatchPress_Interface.bHeatStakeCommissioned,
    bVisionCommissioned := GVL_PatchPress_Interface.bVisionCommissioned,
    bCoreCommissioningMode := GVL_PatchPress_Interface.bCoreCommissioningMode,
    bLogoutHMI := FALSE,
    stOutputs => GVL_MASTER.stOutputs,
    stStatus => GVL_MASTER.stStatus);

END_PROGRAM

// ---- POUs/01_Core/Machine/FB_IndexedPatchPressMachine.TcPOU
FUNCTION_BLOCK FB_IndexedPatchPressMachine
VAR
    fbIndex : FB_IndexTable4;
    fbMainDoorLock : FB_MainDoorLock;
    fbNestManager : FB_NestTableManager;
    fbOperatorStation : FB_OperatorStation;
    fbPatchDispense : FB_PatchDispenseStation;
    fbHeatStake : FB_HeatStakeStation;
    fbVision : FB_VisionStation;
    fbCommissioningGuard : FB_PatchPressCommissioningGuard;
    eMachineState : E_MachineState := E_MachineState.PowerUp;
    eInitialisingWaitReason : E_InitialisingWaitReason := E_InitialisingWaitReason.None;
    eStoppingWaitReason : E_StoppingWaitReason := E_StoppingWaitReason.None;
    stOutputsInternal : ST_MachineOutputs;
    stIndexStatus : ST_IndexStatus;
    stMainDoorStatus : ST_MainDoorLockStatus;
    stOperatorStatus : ST_OperatorStationStatus;
    stPatchDispenseStatus : ST_PatchStageStatus;
    stHeatStakeStatus : ST_PatchStageStatus;
    stVisionStatus : ST_PatchStageStatus;
    stOperatorNest : ST_Nest;
    stPermissives : ST_MachinePermissives;
    tonInitialising : TON;
    tonStopping : TON;
    bInitialisationTimeoutFault : BOOL;
    bStoppingTimeoutFault : BOOL;
    bAutoCycleAllowed : BOOL;
    sAutoCycleBlockReason : STRING(160);
    bIndexMoveAccepted : BOOL;
    bDoorLockOutput : BOOL;
    rtManualIndexMove : R_TRIG;
    rtCoreAutoIndexMove : R_TRIG;
END_VAR

METHOD PUBLIC Cyclic
VAR_INPUT
    stInputs : ST_MachineInputs;
    stCommand : ST_MachineCommand;
    stConfig : ST_MachineConfig;
    bPatchDispenseCommissioned : BOOL;
    bHeatStakeCommissioned : BOOL;
    bVisionCommissioned : BOOL;
    bCoreCommissioningMode : BOOL;
    bLogoutHMI : BOOL;
END_VAR
VAR_OUTPUT
    stOutputs : ST_MachineOutputs;
    stStatus : ST_MachineStatus;
END_VAR
ResetCyclicOutputs();
fbNestManager.Cyclic(bIndexStable := stInputs.bIndexReady AND stInputs.bIndexLocked, eIndexPosition := stInputs.eIndexPosition, eOperatorPosition := stConfig.eOperatorPosition, bPartPresent := stInputs.bLoadingStationEaglePresent, aNestEnabled := stConfig.aNestEnabled);
stOperatorNest := fbNestManager.GetNestAtPosition(stConfig.eOperatorPosition);
fbOperatorStation.Cyclic(bAutomaticActive := (eMachineState = E_MachineState.AutoCycle), bIndexStable := stInputs.bIndexReady AND stInputs.bIndexLocked, stOperatorNest := stOperatorNest, bPartPresent := stInputs.bLoadingStationEaglePresent, bRejectChutePartPresent := stInputs.bRejectChutePartPresent, bRequireRejectConfirm := stConfig.bRequireRejectConfirm, bAllowEmptyNestIndex := stConfig.bAllowEmptyNestIndex);
stOperatorStatus := fbOperatorStation.GetStatus();
fbPatchDispense.Cyclic(bEnable := (eMachineState = E_MachineState.AutoCycle), bCommissioned := bPatchDispenseCommissioned, bStart := FALSE, bReset := stCommand.bReset, bSafetyOk := stInputs.stSafety.bSafetyOk, stStatus => stPatchDispenseStatus);
fbHeatStake.Cyclic(bEnable := (eMachineState = E_MachineState.AutoCycle), bCommissioned := bHeatStakeCommissioned, bStart := FALSE, bReset := stCommand.bReset, bSafetyOk := stInputs.stSafety.bSafetyOk, stStatus => stHeatStakeStatus);
fbVision.Cyclic(bEnable := (eMachineState = E_MachineState.AutoCycle), bCommissioned := bVisionCommissioned, bStart := FALSE, bReset := stCommand.bReset, bSafetyOk := stInputs.stSafety.bSafetyOk, stStatus => stVisionStatus);
stPermissives.bAirSupplyReady := GVL_Safety.bAirSupplySafe;
stPermissives.bDoorInitialisationReady := stInputs.bMainDoorClosed AND NOT stInputs.bMainDoorUnsafe;
stPermissives.bIndexInitialisationReady := NOT fbIndex.IsFaulted();
stPermissives.bStationsHome := TRUE;
stPermissives.bInitialisationAllowed := stInputs.stSafety.bSafetyOk AND stPermissives.bAirSupplyReady AND stPermissives.bDoorInitialisationReady AND stPermissives.bIndexInitialisationReady;
stPermissives.bSafetyIndexPermissive := stInputs.stSafety.bMotionSafetyPermitted;
stPermissives.bOperatorIndexPermissive := stOperatorStatus.bIndexPermissive;
stPermissives.bStationsIndexPermissive := TRUE;
stPermissives.bIndexMoveAllowed := stPermissives.bSafetyIndexPermissive AND stPermissives.bStationsIndexPermissive;
fbCommissioningGuard.Cyclic(bDispenseCommissioned := bPatchDispenseCommissioned, bHeatStakeCommissioned := bHeatStakeCommissioned, bVisionCommissioned := bVisionCommissioned, bCoreCommissioningMode := bCoreCommissioningMode, bCoreReady := ((eMachineState = E_MachineState.ReadyToStart) OR (eMachineState = E_MachineState.AutoCycle)), bAutoCycleAllowed => bAutoCycleAllowed, sBlockReason => sAutoCycleBlockReason);
stPermissives.bAutoCycleAllowed := bAutoCycleAllowed;
IF stInputs.bEventFault OR fbIndex.IsFaulted() OR fbMainDoorLock.IsFaulted() THEN eMachineState := E_MachineState.Fault; END_IF
CASE eMachineState OF
E_MachineState.PowerUp:
    // Same lifecycle used by the validated Silicone Station core:
    // always enter a controlled stop before waiting for Reset.
    tonInitialising(IN := FALSE);
    tonStopping(IN := FALSE);
    eMachineState := E_MachineState.Stopping;

E_MachineState.Stopping:
    tonInitialising(IN := FALSE);
    tonStopping(IN := stIndexStatus.bBusy, PT := stConfig.tStoppingTimeout);
    bStoppingTimeoutFault := tonStopping.Q;
    IF bStoppingTimeoutFault THEN
        eMachineState := E_MachineState.Fault;
    ELSIF NOT stIndexStatus.bBusy THEN
        eMachineState := E_MachineState.Stopped;
    END_IF

E_MachineState.Stopped:
    tonInitialising(IN := FALSE);
    tonStopping(IN := FALSE);
    IF stCommand.bReset AND stInputs.stSafety.bSafetyOk THEN
        eMachineState := E_MachineState.Initialising;
    END_IF

E_MachineState.Initialising:
    stOutputsInternal.bSafetyRunRequest := TRUE;
    stOutputsInternal.bAirSupplyEnable := TRUE;
    tonStopping(IN := FALSE);
    tonInitialising(IN := NOT stPermissives.bInitialisationAllowed, PT := stConfig.tInitialiseTimeout);
    bInitialisationTimeoutFault := tonInitialising.Q;
    IF bInitialisationTimeoutFault THEN
        eMachineState := E_MachineState.Fault;
    ELSIF stPermissives.bInitialisationAllowed THEN
        tonInitialising(IN := FALSE);
        eMachineState := E_MachineState.ReadyToStart;
    END_IF

E_MachineState.ReadyToStart:
    stOutputsInternal.bSafetyRunRequest := TRUE;
    stOutputsInternal.bAirSupplyEnable := TRUE;
    IF stCommand.bStop THEN
        eMachineState := E_MachineState.Stopping;
    ELSIF stCommand.bManualRequest
        AND stInputs.stSafety.bSafetyOk
        AND NOT stIndexStatus.bBusy
        AND NOT fbIndex.IsFaulted()
    THEN
        eMachineState := E_MachineState.Manual;
    ELSIF stCommand.bStart AND bAutoCycleAllowed AND fbMainDoorLock.IsReadyForAutomatic() THEN
        eMachineState := E_MachineState.AutoCycle;
    END_IF

E_MachineState.AutoCycle:
    stOutputsInternal.bSafetyRunRequest := TRUE;
    stOutputsInternal.bAirSupplyEnable := TRUE;
    IF stCommand.bStop OR stInputs.bEventCycleStopRequest THEN
        eMachineState := E_MachineState.Stopping;
    END_IF

E_MachineState.Manual:
    stOutputsInternal.bSafetyRunRequest := TRUE;
    stOutputsInternal.bAirSupplyEnable := TRUE;
    IF stCommand.bStop OR NOT stCommand.bManualRequest THEN
        eMachineState := E_MachineState.Stopping;
    END_IF

E_MachineState.Fault:
    tonInitialising(IN := FALSE);
    tonStopping(IN := FALSE);
    IF stCommand.bReset
        AND NOT stInputs.bEventFault
        AND stInputs.stSafety.bSafetyOk
    THEN
        bInitialisationTimeoutFault := FALSE;
        bStoppingTimeoutFault := FALSE;
        fbIndex.Reset();
        eMachineState := E_MachineState.Stopping;
    END_IF
END_CASE

// Manual Index follows the validated Silicone Station behaviour:
// enable the Indexer on the HMI, then a fresh two-hand actuation requests one move.
rtManualIndexMove(CLK :=
    (eMachineState = E_MachineState.Manual)
    AND stCommand.bIndexerManualEnable
    AND stInputs.bTwoHandsSafe);

IF rtManualIndexMove.Q THEN
    bIndexMoveAccepted := fbIndex.RequestManualMove();
END_IF

// Engineering-only automatic index commissioning. This is deliberately
// isolated from the future production ProcessCycle. Every fresh two-hand
// actuation requests exactly one index step.
rtCoreAutoIndexMove(CLK :=
    (eMachineState = E_MachineState.AutoCycle)
    AND bCoreCommissioningMode
    AND stInputs.bTwoHandsSafe);

IF rtCoreAutoIndexMove.Q THEN
    bIndexMoveAccepted := fbIndex.RequestMove();
END_IF
fbIndex.Cyclic(bEnable := (eMachineState <> E_MachineState.PowerUp) AND (eMachineState <> E_MachineState.Fault), bReset := stCommand.bReset, bAutomaticMode := (eMachineState = E_MachineState.AutoCycle), bManualMode := (eMachineState = E_MachineState.Manual), bMovePermissive := stPermissives.bIndexMoveAllowed, bSafetyMotionPermitted := stInputs.stSafety.bMotionSafetyPermitted, bTwoHandsSafe := stInputs.bTwoHandsSafe, bStationsHome := TRUE, bProcessToolingRetracted := TRUE, bTableReady := stInputs.bIndexReady, bTableLocked := stInputs.bIndexLocked, bCompletedSensor := stInputs.bIndexCompletedSensor, bSupportExtended := TRUE, bSupportRetracted := TRUE, eCurrentPosition := stInputs.eIndexPosition, tRotateDelay := stConfig.tIndexRotateDelay, tStopDelay := stConfig.tIndexStopDelay, tSupportTimeout := stConfig.tIndexSupportTimeout, tMovementTimeout := stConfig.tIndexTimeout, tTwoHandHold := stConfig.tTwoHandHold, tTwoHandRecoveryTimeout := stConfig.tTwoHandRecoveryTimeout, bRotatePortA => stOutputsInternal.bIndexRotatePortA, bStopPortB => stOutputsInternal.bIndexStopPortB, bSupportExtendRequest => stOutputsInternal.bIndexSupportExtend, bSupportRetractRequest => stOutputsInternal.bIndexSupportRetract);
stIndexStatus := fbIndex.GetStatus();
fbMainDoorLock.Cyclic(bEnableAutomatic := (eMachineState = E_MachineState.Initialising) OR (eMachineState = E_MachineState.ReadyToStart) OR (eMachineState = E_MachineState.AutoCycle), bManualEnable := (eMachineState = E_MachineState.Manual), bManualLockRequest := NOT stCommand.bManualMainDoorUnlock, bManualUnlockRequest := stCommand.bManualMainDoorUnlock, bStopRequest := (eMachineState = E_MachineState.Stopping), bResetRequest := stCommand.bReset, bDoorClosed := stInputs.bMainDoorClosed, bDoorLocked := stInputs.bMainDoorLocked, bIndexBusy := stIndexStatus.bBusy, bProcessSafePosition := TRUE, tLockTimeout := stConfig.tDoorLockTimeout, tUnlockTimeout := stConfig.tDoorUnlockTimeout, bDoorUnsafe := stInputs.bMainDoorUnsafe, bLockOutput => bDoorLockOutput);
stOutputsInternal.bMainDoorLockRequest := bDoorLockOutput;
stMainDoorStatus := fbMainDoorLock.GetStatus();
stOutputsInternal.bSafetyResetRequest := stCommand.bReset;
stOutputsInternal.bSafetyErrorAcknowledgementRequest := stCommand.bReset;
stOutputsInternal.bLedStart := (eMachineState = E_MachineState.ReadyToStart);
stOutputsInternal.bLedReset := (eMachineState = E_MachineState.Fault);
stOutputsInternal.bLedPass := (eMachineState = E_MachineState.AutoCycle);
stOutputsInternal.bLedFail := (eMachineState = E_MachineState.Fault);
stOutputsInternal.bInternalLight := TRUE;
stOutputsInternal.bNestLight := TRUE;
stOutputs := stOutputsInternal;
stStatus.eMachineState := eMachineState;
stStatus.eIndexState := fbIndex.GetState();
stStatus.stIndexStatus := stIndexStatus;
stStatus.stMainDoorLock := stMainDoorStatus;
stStatus.eInitialisingWaitReason := eInitialisingWaitReason;
stStatus.eStoppingWaitReason := eStoppingWaitReason;
stStatus.eOperatorExchangeState := fbOperatorStation.GetState();
stStatus.eOperatorInstruction := fbOperatorStation.GetInstruction();
stStatus.stOperatorStation := stOperatorStatus;
stStatus.stPatchDispense := stPatchDispenseStatus;
stStatus.stHeatStake := stHeatStakeStatus;
stStatus.stVision := stVisionStatus;
stStatus.bReady := (eMachineState = E_MachineState.ReadyToStart);
stStatus.bBusy := (eMachineState = E_MachineState.AutoCycle) OR stIndexStatus.bBusy;
stStatus.bFaulted := (eMachineState = E_MachineState.Fault);
stStatus.bInitialisationTimeoutFault := bInitialisationTimeoutFault;
stStatus.bStoppingTimeoutFault := bStoppingTimeoutFault;
stStatus.bSafetyStopRequested := NOT stInputs.stSafety.bSafetyOk;
stStatus.bSafetyRunRequested := stOutputsInternal.bSafetyRunRequest;
stStatus.bEventFault := stInputs.bEventFault;
stStatus.bCycleStopRequested := stInputs.bEventCycleStopRequest;
stStatus.bIndexPermissive := stPermissives.bIndexMoveAllowed;
stStatus.bEnableSetting := (eMachineState = E_MachineState.Stopped) OR (eMachineState = E_MachineState.Manual);
stStatus.bAllStationsCommissioned := bPatchDispenseCommissioned AND bHeatStakeCommissioned AND bVisionCommissioned;
stStatus.bAutoCycleAllowed := bAutoCycleAllowed;
stStatus.stPermissives := stPermissives;
stStatus.aNest := fbNestManager.GetAllNests();
stStatus.aNestStatistics := fbNestManager.GetAllNestStatistics();
stStatus.sAutoCycleBlockReason := sAutoCycleBlockReason;
CASE eMachineState OF
    E_MachineState.PowerUp: stStatus.sMachineMessage := 'System power up';
    E_MachineState.Initialising: stStatus.sMachineMessage := 'System initialising';
    E_MachineState.ReadyToStart: IF bAutoCycleAllowed THEN stStatus.sMachineMessage := 'System ready to start'; ELSE stStatus.sMachineMessage := sAutoCycleBlockReason; END_IF
    E_MachineState.AutoCycle: stStatus.sMachineMessage := 'System auto cycle';
    E_MachineState.Manual: stStatus.sMachineMessage := 'Manual mode';
    E_MachineState.Stopping: stStatus.sMachineMessage := 'Stopping';
    E_MachineState.Stopped: stStatus.sMachineMessage := 'Cycle stopped';
    E_MachineState.Fault: stStatus.sMachineMessage := 'Immediate fault';
END_CASE
END_METHOD

METHOD PRIVATE ResetCyclicOutputs
stOutputsInternal.bSafetyRunRequest := FALSE;
stOutputsInternal.bSafetyResetRequest := FALSE;
stOutputsInternal.bSafetyErrorAcknowledgementRequest := FALSE;
stOutputsInternal.bAirSupplyEnable := FALSE;
stOutputsInternal.bMainDoorLockRequest := FALSE;
stOutputsInternal.bIndexRotatePortA := FALSE;
stOutputsInternal.bIndexStopPortB := FALSE;
stOutputsInternal.bIndexSupportExtend := FALSE;
stOutputsInternal.bIndexSupportRetract := FALSE;
stOutputsInternal.bLedStart := FALSE;
stOutputsInternal.bLedReset := FALSE;
stOutputsInternal.bLedPass := FALSE;
stOutputsInternal.bLedFail := FALSE;
END_METHOD

END_FUNCTION_BLOCK

// ---- POUs/02_Components/Index/FB_IndexTable4.TcPOU
FUNCTION_BLOCK FB_IndexTable4
VAR
    eState                         : E_IndexState := E_IndexState.Initialising;
    eFault                         : E_IndexFault := E_IndexFault.None;
    ePositionAtMoveStart           : E_TablePosition := E_TablePosition.Unknown;
	eStateBeforeWrongPosition       : E_IndexState := E_IndexState.Idle;
	
    bRequestPending                : BOOL;
    bDonePulse                     : BOOL;
    bManualMoveActive              : BOOL;
    bPositionRecoveryActive        : BOOL;
    bWrongPositionSupervisionActive: BOOL;
    bReleaseProcessPosition        : BOOL;
    bOperatorExchangeDone          : BOOL;
	bSamePositionDetected 		   : BOOL;
	
	
    tonTwoHandHold                 : TON;
    tonRotateDelay                 : TON;
    tonStopDelay                   : TON;
    tonStateTimeout                : TON;
    tonWrongPosition               : TON;
	
	
    stInternalStatus               : ST_IndexStatus;
END_VAR

METHOD PUBLIC ConfirmOperatorExchange
IF eState = E_IndexState.WaitingOperatorExchange THEN bOperatorExchangeDone := TRUE; END_IF
END_METHOD

METHOD PUBLIC Cyclic
VAR_INPUT
    bEnable                 : BOOL;
    bReset                  : BOOL;
    bAutomaticMode          : BOOL;
    bManualMode             : BOOL;
    bMovePermissive         : BOOL;
    bSafetyMotionPermitted  : BOOL;
    bTwoHandsSafe           : BOOL;
    bStationsHome           : BOOL;
    bProcessToolingRetracted: BOOL;
    bTableReady             : BOOL;
    bTableLocked            : BOOL;
    bCompletedSensor        : BOOL;
    bSupportExtended        : BOOL;
    bSupportRetracted       : BOOL;
    eCurrentPosition        : E_TablePosition;
    tRotateDelay            : TIME;
    tStopDelay              : TIME;
    tSupportTimeout         : TIME;
    tMovementTimeout        : TIME;
    tTwoHandHold            : TIME;
    tTwoHandRecoveryTimeout : TIME;
END_VAR
VAR_OUTPUT
    bRotatePortA            : BOOL;
    bStopPortB              : BOOL;
    bSupportExtendRequest   : BOOL;
    bSupportRetractRequest  : BOOL;
END_VAR
// =========================================================
// DETERMINISTIC OUTPUT DEFAULTS
// =========================================================

bRotatePortA := FALSE;
bStopPortB := FALSE;

// Support-cylinder outputs are not used during the current commissioning stage.
bSupportExtendRequest := FALSE;
bSupportRetractRequest := FALSE;

bDonePulse := FALSE;


// =========================================================
// TIMERS
// =========================================================

// Temporarily disabled.
//
// The index movement starts immediately when the validated two-hand signal
// becomes TRUE. A minimum hold time is not currently required.
//
// tonTwoHandHold(
//     IN := bTwoHandsSafe,
//     PT := tTwoHandHold
// );

tonRotateDelay(
    IN := eState = E_IndexState.RotatingPortA,
    PT := tRotateDelay
);

tonStopDelay(
    IN := eState = E_IndexState.StoppingPortB,
    PT := tStopDelay
);

tonWrongPosition(
    IN := bWrongPositionSupervisionActive,
    PT := tTwoHandRecoveryTimeout
);


// Only active movement states are supervised during the current
// index commissioning stage.
tonStateTimeout(
    IN :=
        eState = E_IndexState.RotatingPortA
        OR eState = E_IndexState.StoppingPortB
        OR eState = E_IndexState.VerifyingPosition,

    PT := tMovementTimeout
);


// Original support supervision retained for future implementation.
//
// tonStateTimeout(
//     IN := eState = E_IndexState.RetractingSupport
//        OR eState = E_IndexState.WaitingSupportRetracted
//        OR eState = E_IndexState.RotatingPortA
//        OR eState = E_IndexState.StoppingPortB
//        OR eState = E_IndexState.VerifyingPosition
//        OR eState = E_IndexState.ExtendingSupport
//        OR eState = E_IndexState.WaitingSupportExtended,
// 
//     PT := SEL(
//         eState = E_IndexState.RotatingPortA
//         OR eState = E_IndexState.StoppingPortB
//         OR eState = E_IndexState.VerifyingPosition,
//         tSupportTimeout,
//         tMovementTimeout
//     )
// );


// =========================================================
// RESET
// =========================================================

IF bReset THEN

    bRequestPending := FALSE;
    bReleaseProcessPosition := FALSE;
    bOperatorExchangeDone := FALSE;

    bManualMoveActive := FALSE;
    bPositionRecoveryActive := FALSE;
    bWrongPositionSupervisionActive := FALSE;

    eFault := E_IndexFault.None;

    IF bEnable THEN
        eState := E_IndexState.Initialising;
    ELSE
        eState := E_IndexState.Disabled;
    END_IF

END_IF


// =========================================================
// DISABLE HANDLING
// =========================================================

IF NOT bEnable
    AND eState <> E_IndexState.Disabled
THEN
    eState := E_IndexState.Disabled;
END_IF


// =========================================================
// INDEX STATE MACHINE
// =========================================================

CASE eState OF


    // =====================================================
    // DISABLED
    // =====================================================

    E_IndexState.Disabled:

        IF bEnable THEN
            eState := E_IndexState.Initialising;
        END_IF


    // =====================================================
    // INITIALISING
    // =====================================================

    E_IndexState.Initialising:

        // Initialising only prepares the index controller.
        // No automatic movement is performed here.
        IF bEnable
            AND bSafetyMotionPermitted
        THEN
            eState := E_IndexState.Idle;
        END_IF


    // =====================================================
    // IDLE
    // =====================================================

    E_IndexState.Idle:

        // Current commissioning requirements:
        //
        // 1. A movement request is pending.
        // 2. Manual movement is permitted.
        // 3. Motion safety is available.
        // 4. The two-hand signal is active.
        //
        // Support-cylinder feedback is temporarily excluded.
        IF bRequestPending
            AND bMovePermissive

            // Temporarily disabled until the support cylinders
            // are commissioned.
            //
            // AND bStationsHome
            // AND bProcessToolingRetracted

            AND bSafetyMotionPermitted
            AND bTwoHandsSafe
        THEN

            bRequestPending := FALSE;
            ePositionAtMoveStart := eCurrentPosition;

            // Support retraction sequence temporarily bypassed.
            //
            // eState := E_IndexState.RetractingSupport;

            eState := E_IndexState.RotatingPortA;
		
		ELSIF eCurrentPosition = E_TablePosition.Unknown THEN
			
			eState := E_IndexState.WrongPositionRecovery;

        END_IF


    // =====================================================
    // SUPPORT RETRACTION
    // TEMPORARILY NOT USED
    // =====================================================

    E_IndexState.RetractingSupport:

        (*
        bSupportRetractRequest := TRUE;

        IF NOT bSafetyMotionPermitted THEN

            eFault := E_IndexFault.SafetyLostDuringMovement;
            eState := E_IndexState.Fault;

        ELSIF NOT bTableLocked
            AND NOT bTwoHandsSafe
        THEN

            bWrongPositionSupervisionActive := TRUE;
            eState := E_IndexState.WrongPositionRecovery;

        ELSIF bSupportRetracted THEN

            eState := E_IndexState.WaitingSupportRetracted;

        ELSIF tonStateTimeout.Q THEN

            eFault := E_IndexFault.SupportRetractTimeout;
            eState := E_IndexState.Fault;

        END_IF
        *)

        // Temporary bypass.
        eState := E_IndexState.RotatingPortA;


    E_IndexState.WaitingSupportRetracted:

        (*
        bSupportRetractRequest := TRUE;

        IF NOT bTableLocked
            AND NOT bTwoHandsSafe
        THEN

            bWrongPositionSupervisionActive := TRUE;
            eState := E_IndexState.WrongPositionRecovery;

        ELSIF bSupportRetracted THEN

            eState := E_IndexState.RotatingPortA;

        ELSIF tonStateTimeout.Q THEN

            eFault := E_IndexFault.SupportRetractTimeout;
            eState := E_IndexState.Fault;

        END_IF
        *)

        // Temporary bypass.
        eState := E_IndexState.RotatingPortA;


    // =====================================================
    // ROTATE TABLE — PORT A
    // =====================================================

    E_IndexState.RotatingPortA:

        // Support output remains disabled until the cylinder is commissioned.
        //
        // bSupportRetractRequest := TRUE;

        // The two-hand condition must be evaluated first because
        // TwinSAFE may remove bSafetyMotionPermitted immediately when
        // either hand is released.
        IF NOT bTableLocked
            AND NOT bTwoHandsSafe
        THEN

            bWrongPositionSupervisionActive := TRUE;
            eState := E_IndexState.WrongPositionRecovery;


        ELSIF NOT bSafetyMotionPermitted THEN

            eFault := E_IndexFault.SafetyLostDuringMovement;
            eState := E_IndexState.Fault;


        ELSIF NOT bMovePermissive THEN

            eFault := E_IndexFault.MovementPermissiveLost;
            eState := E_IndexState.Fault;


        ELSE

            bRotatePortA := TRUE;

            IF tonRotateDelay.Q
                AND bCompletedSensor
            THEN

                eState := E_IndexState.StoppingPortB;

            ELSIF tonStateTimeout.Q THEN

                eFault := E_IndexFault.RotationTimeout;
                eState := E_IndexState.Fault;

            END_IF

        END_IF


    // =====================================================
    // TWO-HAND RECOVERY
    // =====================================================
	// =====================================================
// TWO-HAND / WRONG-POSITION RECOVERY
// =====================================================
	E_IndexState.WrongPositionRecovery:
	
		// Port B is activated first so that the table can stop
		// and lock safely after the two-hand signal is released.
		bStopPortB := TRUE;
	
	
		// -------------------------------------------------
		// TABLE STOPPED AND LOCKED
		// -------------------------------------------------
		// Once the table is locked, the two-hand command is no
		// longer required. Continue with position verification.
		IF bTableReady
			AND bTableLocked
			AND eCurrentPosition <> E_TablePosition.Unknown
		THEN
	
			bWrongPositionSupervisionActive := FALSE;
			eState := E_IndexState.VerifyingPosition;
		
		ELSIF  bTwoHandsSafe AND eCurrentPosition = E_TablePosition.Unknown THEN
			 bStopPortB := FALSE;
			 bRotatePortA := TRUE;
		
			IF tonRotateDelay.Q
				AND bCompletedSensor THEN
				
				eState := E_IndexState.StoppingPortB;
			END_IF
		// -------------------------------------------------
		// RECOVERY TIMEOUT
		// -------------------------------------------------
		ELSIF tonWrongPosition.Q THEN
	
			bWrongPositionSupervisionActive := FALSE;
	
			eFault := E_IndexFault.WrongPositionTimeout;
			eState := E_IndexState.Fault;
	
	
		// -------------------------------------------------
		// OPERATOR RESTORED BOTH HANDS BEFORE TABLE LOCKED
		// -------------------------------------------------
		ELSIF bTwoHandsSafe
			AND bSafetyMotionPermitted
			AND bMovePermissive
			AND bTableLocked
		THEN
	
			bWrongPositionSupervisionActive := FALSE;
	
			// Resume the exact state interrupted by the
			// two-hand signal release.
			eState := eStateBeforeWrongPosition;
	
		END_IF
    // =====================================================
    // STOP TABLE — PORT B
    // =====================================================

    E_IndexState.StoppingPortB:

        // Support output temporarily disabled.
        //
        // bSupportRetractRequest := TRUE;

        // Continue requiring two hands until the table is locked.
        // This check must be evaluated before bSafetyMotionPermitted.
        IF NOT bTableLocked
            AND NOT bTwoHandsSafe
        THEN

            bWrongPositionSupervisionActive := TRUE;
            eState := E_IndexState.WrongPositionRecovery;


        ELSIF NOT bSafetyMotionPermitted THEN

            eFault := E_IndexFault.SafetyLostDuringMovement;
            eState := E_IndexState.Fault;


        ELSE

            bStopPortB := TRUE;

            IF tonStopDelay.Q
                AND bTableReady
                AND bTableLocked
            THEN

                eState := E_IndexState.VerifyingPosition;

            ELSIF tonStateTimeout.Q THEN

                eFault := E_IndexFault.StopAndLockTimeout;
                eState := E_IndexState.Fault;

            END_IF

        END_IF


    // =====================================================
	// VERIFY NEW POSITION
	// =====================================================
	E_IndexState.VerifyingPosition:
	
		// Support output temporarily disabled.
		//
		// bSupportRetractRequest := TRUE;
	
	
		// At this point the table is already confirmed ready and locked.
		// Two hands are therefore no longer required.
	
		IF eCurrentPosition = E_TablePosition.Unknown THEN
	
			IF tonStateTimeout.Q THEN
	
				eFault := E_IndexFault.PositionInvalid;
				//eState := E_IndexState.Fault;
	
			END_IF
	
	
		ELSIF NOT bPositionRecoveryActive
			AND eCurrentPosition = ePositionAtMoveStart
		THEN
	
			// A valid and known position was detected, but it is the
			// same position from which the movement started.
			//
			// This is process information only and is not an index fault.
			bSamePositionDetected := TRUE;
	
			bWrongPositionSupervisionActive := FALSE;
			eState := E_IndexState.Complete;
	
	
		ELSE
	
			bSamePositionDetected := FALSE;
			bWrongPositionSupervisionActive := FALSE;
	
			// Support extension sequence temporarily bypassed.
			//
			// eState := E_IndexState.ExtendingSupport;
	
			eState := E_IndexState.Complete;
	
		END_IF


    // =====================================================
    // SUPPORT EXTENSION
    // TEMPORARILY NOT USED
    // =====================================================

    E_IndexState.ExtendingSupport:

        (*
        bSupportExtendRequest := TRUE;

        IF bSupportExtended THEN

            eState := E_IndexState.WaitingSupportExtended;

        ELSIF tonStateTimeout.Q THEN

            eFault := E_IndexFault.SupportExtendTimeout;
            eState := E_IndexState.Fault;

        END_IF
        *)

